(* IEC 61131-3 sources: daoli-st-library/DL_Process (part 61) *)

(* ---- FB_DL_BatchDosingControl.st ---- *)
(*==============================================================================
 * 组件名称 (Component)  : FB_DL_BatchDosingControl
 * 所属子库 (Sublibrary) : DL_Process
 * 当前版本 (Version)    : 1.0.1
 * 兼容性 (Platform)   : CODESYS 3.5 / TwinCAT 3 / 汇川 InoProShop / Machine Expert
 *                         仅依赖 Standard.library（TON / R_TRIG），零厂商方言
 * 分类     (Category)   : 工艺功能块（Function Block · 多原料单通道配料称重）
 * 功能简述 (Function)   : 多原料单通道自动配料称重控制器（单料批次相 Phase
 *                         语义）。三段给料顺控（快加→慢加→落定结算）+ 空中
 *                         落差自学习（误差/2 更新，防振荡）+ 超差 NG 判定 +
 *                         断流诊断。执行机构抽象为三离散输出（与给料机/闸门
 *                         类型解耦）；秤重量 LREAL→REAL 引脚注入（标定由称
 *                         重层完成）。Abort 优先级最高（CASE 首分支）。
 * 枚举归属 (Enum note)  : E_DL_DosingPhase 随本块同文件发布（公约 0.11 口径：
 *                         配套枚举与主块同文件，头注释注明归属）。
 * 公约遵循 (Convention) : 0.1/R23 显式批次启动沿驱动（无自动首扫初始化语义），
 *                         免首扫，无 bInit。
 *                         0.2/R21 bFault 显式排除信息级码；0.5/R7 全部实例主
 *                         体最前部无条件刷新；0.7/R15 断流/秤信号/参数故障锁
 *                         存仅复位路径清码；0.9 非有限值 fWeight 防御（自比
 *                         检测，故障级中止全断）；0.14 全部除法/浮点判等走
 *                         ABS 容差。
 *                         0.8 故障码段位 16#0005_xxxx（经 DL_Process
 *                         VERSION.md 码表核对，0005_0220~0223 / 0005_0114~0106
 *                         均未占用）：
 *                         【故障级】0005_0220 断流/堵料、0005_0221 秤信号无
 *                         效（非有限值）、0005_0223 配方参数非法、0005_0222
 *                         非法状态兜底；
 *                         【信息级】0005_0114 稳窗超时按当前值结算、0005_0115
 *                         补偿学习触限。
 * 红线自检 (Redline)    : R1 零全局变量表/外部变量引用 ✓｜R2 零物理 IO 地址 ✓
 *                         R3 纯 IEC 61131-3 ✓｜R4 非有限值中止全断/防振荡半
 *                         误差学习/限幅钳位 ✓
 *                         R5 全变量中英双语同行注释 ✓｜R6 ENUM+CASE+ELSE，Abort
 *                         首分支最高优先 ✓
 *                         R7 五实例（R_TRIG×3/TON×2）主体最前部无条件刷新 ✓
 *                         R8 全常量化 ✓
 * 设计要点 (Key notes)  : ① 截断点公式：慢加关断重量 = fSetpoint −
 *                           fInflightComp；fInflightComp 初值 0 → 首批必然过
 *                           冲 → 学习链收敛（首批预期在注释写明）；
 *                         ② 自学习更新：结算后 Error = fFinalWeight −
 *                           fSetpoint；bLearnEnable 时 fInflightComp +=
 *                           Error/2.0（半误差防振荡），钳位 ±fCompLimit，
 *                           触限置信息级 0005_0115；
 *                         ③ 稳窗判稳：tSettleWindow 内重量变化 <
 *                           fFlowDeadband 才结算；超窗未稳重试
 *                           DL_SETTLE_RETRY_MAX 次后按当前值结算 + 信息级；
 *                         ④ 断流诊断：给料相中 tFlowWatch 窗内重量变化 <
 *                           fFlowDeadband → 断流故障锁存（快加/慢加独立监
 *                           视计时重启）；
 *                         ⑤ 超差 NG 锁存 + 卸料输出禁止（NG 不得流入下工
 *                           序）；Abort 电平最高优先（CASE 首分支，立即关全
 *                           部输出）；
 *                         ⑥ 非有限值 fWeight → 批次中止故障级 0005_0221，
 *                           输出全断。
 * 偏离留档 (Deviation)  : 依 R11 头注释留档，共 1 条：
 *                         ① 新增故障码 0005_0223 配方参数非法：规格故障集未
 *                           覆盖 fSetpoint/fTolerance 非法值路径，编码时补
 *                           充登记（核对 DL_Process 码表未占用）。
 * 开源溯源 (Origin)     : 来源标签 lbp-batch-dosing / isa-88（RAW_NOTES_R7
 *                         S-10：ISA-88 批次相（Phase）语义与重力失重式/增
 *                         量式配料公开工程惯例——三段给料、空中落差补偿、
 *                         半误差学习（提取点②③⑤），公开技术资料，仅借鉴
 *                         语义域；状态机、学习与诊断实现、码位与引脚契约
 *                         100% 本库独立设计，clean-room 未复制源码）。
 * 验收向量 (Acceptance) :
 *   V1 三段给料逐拍：快加至 fSetpoint−fInflightComp 切慢加，同点关断进落定；
 *   V2 学习链 5 批收敛数值复算：首批过冲 Δ → 补偿 +Δ/2 → 逐批 Δ 减半；
 *   V3 补偿限幅：学习值触及 ±fCompLimit → 信息级 0005_0115；
 *   V4 断流：给料中 tFlowWatch 内重量变化 < fFlowDeadband → 0005_0220；
 *   V5 超差 NG + 卸料禁止：|误差| > fTolerance → eNg、bOutDischarge=FALSE；
 *   V6 中止优先级：任意相 bCmdAbort 电平 → 全输出断进 eAbort；
 *   V7 非有限值注入：fWeight=NaN → 0005_0221 输出全断。
 * 修订历史 (Revision)   :
 *   2026-11-15  v1.0.0  首版入库（Round 07 · DL_Process 配料称重件）
 *   2026-11-15  v1.0.1  终审修复 2 处：① _bSettleRestart/_bFlowRestart 单拍
 *                       重启标志永不自清 → 稳窗 TON 永久失效（eSettling 永
 *                       久挂起、判稳拍结算死锁）+ 断流诊断一次后失效（段 1
 *                       实例调用后自清，R24 同源范式）；② fTareOffset/
 *                       fInflightComp 缺 0.9 非数防御（NaN 扩散进净重/截
 *                       断点链路），新增 _fTareEff/_fCompEff 生效值
 *============================================================================*)

(*-----------------------------------------------------------------------------
 * 枚举: E_DL_DosingPhase（归属 FB_DL_BatchDosingControl，与其同文件）
 * 含义: 单料批次相离散状态。编号步长 10 留空位，eFault 取 99 保证排序末位
 *       （全库枚举编号惯例）。
 *----------------------------------------------------------------------------*)
TYPE E_DL_DosingPhase :
(
    eIdle     := 0,   // 空闲：等待批次启动 / Idle, awaiting batch start
    eCoarse   := 10,  // 快加：粗给料输出有效 / Coarse feed active
    eFine     := 20,  // 慢加：细给料输出有效 / Fine feed active
    eSettling := 30,  // 落定：稳窗判稳中 / Settling, stability window judging
    eDone     := 40,  // 完成：批次合格，卸料输出有效 / Done, batch OK, discharge active
    eNg       := 50,  // 超差：批次 NG 锁存，卸料禁止 / NG latched, discharge forbidden
    eAbort    := 60,  // 中止：Abort 电平保持中，全输出断 / Aborted, all outputs off
    eFault    := 99   // 故障锁存：断流/秤信号/参数非法/非法状态 / Latched fault
) UINT;
END_TYPE

FUNCTION_BLOCK FB_DL_BatchDosingControl
VAR_INPUT
    bCmdBatchStart : BOOL;              // 批次启动指令（Batch start），上升沿进入快加 / Batch start edge enters coarse feed
    bCmdAbort      : BOOL;              // 批次中止指令（Abort），电平生效，立即关全部输出 / Abort level, all outputs off immediately
    fWeight        : REAL;              // 秤实时重量（Live weight）[kg]，非有限值防御；标定由称重层完成 / Live weight [kg], non-finite defended, calibration upstream
    fTareOffset    : REAL := 0.0;       // 皮重偏移（Tare offset）[kg]，默认 0.0；净重 = fWeight − fTareOffset / Tare offset [kg], net = weight − tare
    fSetpoint      : REAL;              // 批次目标净重（Batch setpoint）[kg]，域 >0 / Batch setpoint [kg], > 0
    fSwitchCoarse  : REAL := 0.0;       // 快加切换点（Coarse-to-fine switch）[kg]，0=默认 85% 设定值（引脚覆盖语义见头注释）/ Coarse switch point, 0 = default 85% of setpoint
    fInflightComp  : REAL;              // 空中落差补偿（In-flight compensation）[kg]，学习值跨批次保持；上下限由 fCompLimit 钳位 / In-flight compensation [kg], learned value clamped by fCompLimit
    fCompLimit     : REAL := 0.0;       // 补偿学习限幅（Compensation limit）[kg]，0=默认 10% 设定值 / Compensation clamp, 0 = default 10% of setpoint
    bLearnEnable   : BOOL;              // 落差自学习使能（Learning enable），TRUE=每批结算后按误差/2 更新 / Learning enable, update by error/2 after each settle
    tSettleWindow  : TIME := T#1S;     // 落定稳窗（Settle window），默认 T#1S，域 500MS~5S 越界钳位 / Settle window, clamped 500MS..5S
    fTolerance     : REAL := 0.0;       // 批次公差（Batch tolerance）[kg]，0=默认 0.5% 设定值语义（引脚显式覆盖）/ Batch tolerance, 0 = default 0.5% of setpoint
    tFlowWatch     : TIME := T#10S;    // 断流监视窗（Flow watchdog），默认 T#10S；给料中重量变化率恒零超窗 → 断流 / Flow watchdog, constant-weight over window = no flow
    fFlowDeadband  : REAL := 0.05;     // 断流判据死区（Flow deadband）[kg]，默认 0.05；稳窗内重量变化 < 死区判断流 / Flow deadband [kg], change below deadband = no flow
    bReset         : BOOL;              // 上升沿复位故障（Reset edge）/ Rising edge resets fault
END_VAR
VAR_OUTPUT
    bOutCoarse    : BOOL;               // 快加输出（Coarse feed output），给料机/闸门快加速率 / Coarse feed output
    bOutFine      : BOOL;               // 慢加输出（Fine feed output）/ Fine feed output
    bOutDischarge : BOOL;               // 卸料输出（Discharge output），批次合格后放料 / Discharge output, opens after batch OK
    fNetWeight    : REAL;               // 当前净重（Net weight）[kg] / Current net weight [kg]
    fFinalWeight  : REAL;               // 上批次结算净重（Final weight）[kg]，落定后锁存 / Final settled weight [kg], latched after settle
    bBatchOk      : BOOL;               // 批次合格（Batch OK），|结算净重 − 设定值| ≤ 公差 / Batch OK verdict
    bFault        : BOOL;               // 故障标志（Fault flag），显式排除信息级 / Fault flag, info codes excluded
    uErrorId      : UDINT;              // 故障码（Error code），16#0005_xxxx 段，0=无故障 / Error code, family 16#0005_xxxx
END_VAR
VAR
    _ePhase        : E_DL_DosingPhase := E_DL_DosingPhase.eIdle; // 内部批次相（Internal dosing phase），属性只读 / Internal phase, read-only via property
    _bFaultLatch   : BOOL;              // 故障锁存标志（Fault latch flag），仅复位路径清除 / Fault latch, cleared only via reset path
    _uErrorIdInt   : UDINT;             // 内部故障级码寄存（Internal fault-level register）/ Internal fault-level register
    _uInfoCode     : UDINT;             // 本拍信息级码（Info code this cycle），瞬时型每拍重算 / Transient info code, recomputed each scan
    _bWeightValid  : BOOL;              // 秤信号有效（Weight signal valid，非有限值防御）/ Weight signal valid flag
    _fNetInt       : REAL;              // 内部净重（Internal net weight）[kg] / Internal net weight [kg]
    _fSetEff       : REAL;              // 防御后生效设定值（Sanitized setpoint）[kg] / Sanitized setpoint [kg]
    _fTolEff       : REAL;              // 防御后生效公差（Sanitized tolerance）[kg] / Sanitized tolerance [kg]
    _fSwitchEff    : REAL;              // 防御后生效快加切换点（Sanitized coarse switch）[kg] / Sanitized coarse switch [kg]
    _fCompLimEff   : REAL;              // 防御后生效补偿限幅（Sanitized compensation clamp）[kg] / Sanitized compensation clamp [kg]
    _fTareEff      : REAL;              // 防御后生效皮重偏移（Sanitized tare offset）[kg]，0.9 非数防御 / Sanitized tare offset [kg] (v1.0.1)
    _fCompEff      : REAL;              // 防御后生效落差补偿（Sanitized in-flight comp）[kg]，0.9 非数防御 / Sanitized in-flight comp [kg] (v1.0.1)
    _fCutCoarse    : REAL;              // 快加→慢加切换重量（Coarse-to-fine cut weight）[kg] / Coarse-to-fine cut weight [kg]
    _fCutFine      : REAL;              // 慢加关断重量（Fine cut weight）[kg]，= 设定值 − 落差补偿 / Fine cut weight [kg]
    _fSettleRef    : REAL;              // 稳窗基准重量（Settle reference weight）[kg] / Settle reference weight [kg]
    _nSettleRetry  : USINT;             // 稳窗重试计数（Settle retry counter）/ Settle retry counter
    _bSettleRestart: BOOL;              // 稳窗重启单拍（Settle restart one-shot）/ Settle restart one-shot
    _fFlowRef      : REAL;              // 断流监视基准重量（Flow-watch reference weight）[kg] / Flow-watch reference weight [kg]
    _bFlowRestart  : BOOL;              // 断流监视重启单拍（Flow-watch restart one-shot）/ Flow-watch restart one-shot
    _bBatchStartEdge : BOOL;            // 批次启动沿（Batch start edge this scan）/ Batch start edge this scan
    _fbTrigStart   : R_TRIG;            // 批次启动沿检测（Batch start edge detector）/ Batch start edge detector
    _fbTrigReset   : R_TRIG;            // 复位沿检测（Reset edge detector）/ Reset edge detector
    _fbTrigAbort   : R_TRIG;            // 中止沿检测（Abort edge detector），沿置中止态（电平保持由段内判定）/ Abort edge detector
    _fbTonSettle   : TON;               // 落定稳窗定时器（Settle window timer）/ Settle window timer
    _fbTonFlow     : TON;               // 断流监视窗定时器（Flow watchdog timer）/ Flow watchdog timer
END_VAR
VAR CONSTANT
    DL_COARSE_FRAC    : REAL := 0.85;   // 快加切换默认比例（Coarse switch default fraction of setpoint）/ Coarse switch default fraction
    DL_COMP_FRAC      : REAL := 0.10;   // 补偿限幅默认比例（Compensation clamp default fraction）/ Compensation clamp default fraction
    DL_TOL_FRAC       : REAL := 0.005;  // 公差默认比例（Tolerance default fraction of setpoint）/ Tolerance default fraction
    DL_LEARN_DIV      : REAL := 2.0;    // 学习半误差除数（Learning half-error divisor），防振荡 / Learning half-error divisor, anti-oscillation
    DL_SETTLE_WIN_MIN : TIME := T#500MS; // 稳窗下限（Settle window lower clamp）/ Settle window lower clamp
    DL_SETTLE_WIN_MAX : TIME := T#5S;   // 稳窗上限（Settle window upper clamp）/ Settle window upper clamp
    DL_SETTLE_RETRY_MAX : USINT := 3;   // 稳窗重试上限（Settle retry max），超限按当前值结算 / Settle retry max, settle as-is beyond
    DL_REAL_EPS       : REAL := 1.0E-6; // 浮点防零容差（Float divide-guard epsilon）/ Float divide-guard epsilon
END_VAR

// ============================================================================
// 段 1｜实例无条件周期刷新（R7/0.5：严禁置于 IF/CASE 分支内）
//      Unconditional per-cycle refresh of all instances (R7/0.5)
// ============================================================================
_fbTrigStart(CLK := bCmdBatchStart);
_fbTrigReset(CLK := bReset);
_fbTrigAbort(CLK := bCmdAbort);
_bBatchStartEdge := _fbTrigStart.Q;   // 本拍启动沿（Start edge this scan）
_fbTonSettle(IN := (_ePhase = E_DL_DosingPhase.eSettling) AND (NOT _bSettleRestart) AND (NOT _bFaultLatch), PT := tSettleWindow); // 稳窗（Settle window）
_fbTonFlow(IN := ((_ePhase = E_DL_DosingPhase.eCoarse) OR (_ePhase = E_DL_DosingPhase.eFine))
           AND (NOT _bFlowRestart) AND (NOT _bFaultLatch), PT := tFlowWatch); // 断流监视窗（Flow watchdog）
// R24 同源范式：单拍重启标志在实例调用之后自清（v1.0.1 修复：原永不自清 →
// 稳窗 TON 永久失效（eSettling 永久挂起、判稳拍结算死锁）+ 断流诊断一次后
// 永久失效）/ One-shot restart flags self-cleared AFTER the instance calls
// (v1.0.1 fix: flags were never cleared, permanently disabling both timers)
_bSettleRestart := FALSE;         // 稳窗重启单拍自清（Settle restart flag self-cleared）
_bFlowRestart := FALSE;           // 断流监视重启单拍自清（Flow restart flag self-cleared）

// ============================================================================
// 段 2｜秤信号防御（0.9）+ 信息级预清零 + 复位路径（R15）
//      Weight sanitation (0.9) + info preset + reset path (R15)
// ============================================================================
_uInfoCode := 0;                  // 信息级瞬时型每拍重算（Transient info recomputed each scan）

IF fWeight <> fWeight THEN        // 非数自比检测（NaN self-compare）
    _bWeightValid := FALSE;       // 秤信号无效（Weight invalid）
    IF _bFaultLatch = FALSE THEN
        _bFaultLatch := TRUE;     // 秤信号无效故障锁存（Invalid weight latch）
        _uErrorIdInt := 16#0005_0221; // 0005_0221 秤信号无效【故障级】/ Invalid weight signal, fault level
        _ePhase := E_DL_DosingPhase.eFault; // 批次中止进故障态（Batch aborted to fault）
    END_IF
ELSE
    _bWeightValid := TRUE;        // 秤信号有效（Weight valid）
    _fNetInt := fWeight - _fTareEff; // 净重计算（皮重经 0.9 非数防御生效值，v1.0.1）/ Net weight with sanitized tare (v1.0.1)
END_IF
fNetWeight := _fNetInt;           // 净重出口（Net weight outlet）

IF _fbTrigReset.Q THEN
    _bFaultLatch := FALSE;        // 故障锁存解除（Fault latch released）
    _uErrorIdInt := 16#0000_0000; // 故障码清零（Fault code cleared）
    IF _ePhase = E_DL_DosingPhase.eFault THEN
        _ePhase := E_DL_DosingPhase.eIdle; // 故障复位回空闲（Fault reset to idle）
    END_IF
END_IF

// ============================================================================
// 段 3｜参数防御（启动时校验配方，0.9 + 域防御）
//      Recipe parameter sanitation at batch start (0.9 + domain guards)
// ============================================================================
IF fSetpoint <> fSetpoint THEN    // 设定值非数（Setpoint NaN）
    _fSetEff := 0.0;              // 非法设定占位（Invalid placeholder）
ELSIF fSetpoint <= DL_REAL_EPS THEN
    _fSetEff := 0.0;              // 非正设定占位（Non-positive placeholder）
ELSE
    _fSetEff := fSetpoint;        // 生效设定（Effective setpoint）
END_IF

IF fTolerance <> fTolerance THEN  // 公差非数（Tolerance NaN）
    _fTolEff := _fSetEff * DL_TOL_FRAC; // 回落默认比例（Default fraction fallback）
ELSIF fTolerance <= 0.0 THEN
    _fTolEff := _fSetEff * DL_TOL_FRAC; // 非正回落默认（Non-positive falls back）
ELSE
    _fTolEff := fTolerance;       // 生效公差（Effective tolerance）
END_IF

IF fSwitchCoarse <> fSwitchCoarse THEN // 切换点非数（Switch NaN）
    _fSwitchEff := _fSetEff * DL_COARSE_FRAC; // 回落默认比例（Default fraction fallback）
ELSIF fSwitchCoarse <= 0.0 THEN
    _fSwitchEff := _fSetEff * DL_COARSE_FRAC; // 零值=默认 85% 设定值（Zero = default 85%）
ELSE
    _fSwitchEff := fSwitchCoarse; // 引脚覆盖生效（Pin override effective）
END_IF

IF fCompLimit <> fCompLimit THEN  // 限幅非数（Clamp NaN）
    _fCompLimEff := _fSetEff * DL_COMP_FRAC; // 回落默认比例（Default fraction fallback）
ELSIF fCompLimit <= 0.0 THEN
    _fCompLimEff := _fSetEff * DL_COMP_FRAC; // 零值=默认 10% 设定值（Zero = default 10%）
ELSE
    _fCompLimEff := fCompLimit;   // 生效限幅（Effective clamp）
END_IF

// 0.9 非数防御补齐（v1.0.1）：皮重偏移与落差补偿为 REAL 输入，非数自比后
// 取生效值，杜绝 NaN 扩散进净重/截断点链路
// 0.9 NaN defense completed (v1.0.1) for tare offset and in-flight compensation
IF fTareOffset <> fTareOffset THEN // 皮重非数（Tare NaN）
    _fTareEff := 0.0;             // 回落零皮重（Fallback zero tare）
ELSE
    _fTareEff := fTareOffset;     // 生效皮重（Effective tare）
END_IF
IF fInflightComp <> fInflightComp THEN // 落差补偿非数（In-flight comp NaN）
    _fCompEff := 0.0;             // 回落零补偿（首批过冲语义，学习链重建）/ Fallback zero comp
ELSE
    _fCompEff := fInflightComp;   // 生效补偿（Effective compensation）
END_IF

// ============================================================================
// 段 4｜主批次相状态机（ENUM + CASE + ELSE 兜底；Abort 首分支最高优先）
//      Main dosing phase machine (Abort first-branch top priority, ELSE fallback)
// ============================================================================
IF bCmdAbort THEN
    // Abort 电平最高优先：立即关全部输出进中止态（Abort level top priority）
    _ePhase := E_DL_DosingPhase.eAbort; // 进中止态（To aborted state）
ELSE
    CASE _ePhase OF

        E_DL_DosingPhase.eIdle: // 空闲态：等待启动沿
            IF _bBatchStartEdge AND (NOT _bFaultLatch) THEN
                IF _fSetEff <= DL_REAL_EPS THEN
                    _bFaultLatch := TRUE;           // 配方参数非法锁存（Invalid recipe latch）
                    _uErrorIdInt := 16#0005_0223;   // 0005_0223 配方参数非法【故障级】/ Invalid recipe parameters, fault level
                    _ePhase := E_DL_DosingPhase.eFault;
                ELSE
                    _fCutCoarse := _fSwitchEff;                     // 快加切换点（Coarse cut point）
                    _fCutFine := _fSetEff - _fCompEff;              // 慢加关断重量 = 设定值 − 落差补偿（截断点公式，生效值）/ Fine cut = setpoint − sanitized comp
                    fFinalWeight := 0.0;                            // 上批结果清位（Final weight cleared）
                    bBatchOk := FALSE;                              // 合格判定清位（OK verdict cleared）
                    _nSettleRetry := 0;                             // 稳窗重试清零（Retry cleared）
                    _fSettleRef := _fNetInt;                        // 稳窗基准初始化（Settle reference init）
                    _fFlowRef := _fNetInt;                          // 断流基准初始化（Flow reference init）
                    _ePhase := E_DL_DosingPhase.eCoarse;            // 进入快加（To coarse feed）
                END_IF
            END_IF

        E_DL_DosingPhase.eCoarse: // 快加态：粗给料至切换点
            IF _fNetInt >= _fCutCoarse THEN
                _ePhase := E_DL_DosingPhase.eFine; // 切慢加（To fine feed）
                _fFlowRef := _fNetInt;             // 断流基准重置（Flow reference reset）
            END_IF

        E_DL_DosingPhase.eFine: // 慢加态：细给料至截断点
            IF _fNetInt >= _fCutFine THEN
                _ePhase := E_DL_DosingPhase.eSettling; // 关断进落定（Cut to settling）
                _fSettleRef := _fNetInt;               // 稳窗基准重置（Settle reference reset）
            END_IF

        E_DL_DosingPhase.eSettling: // 落定态：稳窗判稳，判稳即一次性结算+学习
            IF _fbTonSettle.Q THEN
                IF ABS(_fNetInt - _fSettleRef) < fFlowDeadband THEN
                    // —— 一次性结算（仅判稳拍执行）：锁存结果 + NG 判定 + 学习 ——
                    //     One-shot settlement on the settled scan: result latch, NG verdict, learning
                    fFinalWeight := _fNetInt;   // 结算净重锁存（Final weight latched）
                    bBatchOk := ABS(fFinalWeight - _fSetEff) <= _fTolEff; // 公差判定（Tolerance verdict）
                    IF bLearnEnable THEN
                        fInflightComp := fInflightComp + (fFinalWeight - _fSetEff) / DL_LEARN_DIV; // 误差/2 学习（半误差防振荡）/ Half-error learning, anti-oscillation
                        IF fInflightComp > _fCompLimEff THEN
                            fInflightComp := _fCompLimEff;  // 正向限幅（Positive clamp）
                            _uInfoCode := 16#0005_0115;     // 0005_0115 补偿学习触限【信息级】/ Learning clamp hit, info level
                        ELSIF fInflightComp < (-_fCompLimEff) THEN
                            fInflightComp := -_fCompLimEff; // 负向限幅（Negative clamp）
                            _uInfoCode := 16#0005_0115;     // 0005_0115 补偿学习触限【信息级】/ Learning clamp hit, info level
                        END_IF
                    END_IF
                    IF bBatchOk THEN
                        _ePhase := E_DL_DosingPhase.eDone;  // 合格进完成态（OK to done）
                    ELSE
                        _ePhase := E_DL_DosingPhase.eNg;    // 超差进 NG 锁存态（Out of tolerance to NG）
                    END_IF
                ELSE
                    _nSettleRetry := _nSettleRetry + 1; // 未稳重试（Retry when unstable）
                    IF _nSettleRetry >= DL_SETTLE_RETRY_MAX THEN
                        _uInfoCode := 16#0005_0114;     // 0005_0114 稳窗超时按当前值结算【信息级】/ Settle timeout, settle as-is, info level
                        fFinalWeight := _fNetInt;       // 按当前值结算锁存（Settle as-is latch）
                        bBatchOk := ABS(fFinalWeight - _fSetEff) <= _fTolEff; // 公差判定（Tolerance verdict）
                        IF bBatchOk THEN
                            _ePhase := E_DL_DosingPhase.eDone;
                        ELSE
                            _ePhase := E_DL_DosingPhase.eNg;
                        END_IF
                    ELSE
                        _fSettleRef := _fNetInt;        // 重置稳窗基准（Reset settle reference）
                        _bSettleRestart := TRUE;        // 稳窗重启单拍（Restart window one-shot）
                    END_IF
                END_IF
            END_IF

        E_DL_DosingPhase.eDone: // 完成态：卸料保持，等待新批次启动
            IF _bBatchStartEdge AND (NOT _bFaultLatch) THEN
                IF _fSetEff <= DL_REAL_EPS THEN
                    _bFaultLatch := TRUE;               // 配方参数非法锁存（Invalid recipe latch）
                    _uErrorIdInt := 16#0005_0223;       // 0005_0223 配方参数非法【故障级】/ Invalid recipe, fault level
                    _ePhase := E_DL_DosingPhase.eFault;
                ELSE
                    _fCutCoarse := _fSwitchEff;         // 快加切换点（Coarse cut point）
                    _fCutFine := _fSetEff - _fCompEff;  // 截断点更新（Fine cut update, sanitized comp）
                    fFinalWeight := 0.0;                // 上批结果清位（Final weight cleared）
                    bBatchOk := FALSE;                  // 合格判定清位（OK verdict cleared）
                    _nSettleRetry := 0;                 // 稳窗重试清零（Retry cleared）
                    _fSettleRef := _fNetInt;            // 稳窗基准初始化（Settle reference init）
                    _fFlowRef := _fNetInt;              // 断流基准初始化（Flow reference init）
                    _ePhase := E_DL_DosingPhase.eCoarse; // 进入快加（To coarse feed）
                END_IF
            END_IF

        E_DL_DosingPhase.eNg: // 超差态：卸料禁止，等待新批次启动或 Abort
            IF _bBatchStartEdge AND (NOT _bFaultLatch) THEN
                IF _fSetEff <= DL_REAL_EPS THEN
                    _bFaultLatch := TRUE;               // 配方参数非法锁存（Invalid recipe latch）
                    _uErrorIdInt := 16#0005_0223;       // 0005_0223 配方参数非法【故障级】/ Invalid recipe, fault level
                    _ePhase := E_DL_DosingPhase.eFault;
                ELSE
                    _fCutCoarse := _fSwitchEff;         // 快加切换点（Coarse cut point）
                    _fCutFine := _fSetEff - _fCompEff;  // 截断点更新（Fine cut update, sanitized comp）
                    fFinalWeight := 0.0;                // 上批结果清位（Final weight cleared）
                    bBatchOk := FALSE;                  // 合格判定清位（OK verdict cleared）
                    _nSettleRetry := 0;                 // 稳窗重试清零（Retry cleared）
                    _fSettleRef := _fNetInt;            // 稳窗基准初始化（Settle reference init）
                    _fFlowRef := _fNetInt;              // 断流基准初始化（Flow reference init）
                    _ePhase := E_DL_DosingPhase.eCoarse; // 重开新批（New batch from coarse）
                END_IF
            END_IF

        E_DL_DosingPhase.eAbort: // 中止态：Abort 电平撤销后回空闲
            IF NOT bCmdAbort THEN
                _ePhase := E_DL_DosingPhase.eIdle; // 电平撤销回空闲（Level dropped, back to idle）
            END_IF

        E_DL_DosingPhase.eFault: // 故障锁存态：复位路径见段 2
            // 等待复位（Await reset）

        ELSE
            // 非法状态兜底：任何越界枚举值强制锁存故障（Illegal state fallback）
            _bFaultLatch := TRUE;           // 故障锁存（Fault latch）
            _uErrorIdInt := 16#0005_0222;   // 0005_0222 非法状态兜底【故障级】/ Illegal state, fault level
            _ePhase := E_DL_DosingPhase.eFault;
    END_CASE
END_IF

// ============================================================================
// 段 5｜输出推导 + 断流诊断 + 输出全断出口断言
//      Output derivation + no-flow diagnosis + all-off exit assertion
// ============================================================================
bOutCoarse := (_ePhase = E_DL_DosingPhase.eCoarse) AND _bWeightValid AND (NOT _bFaultLatch); // 快加输出派生（Coarse derived form）
bOutFine := (_ePhase = E_DL_DosingPhase.eFine) AND _bWeightValid AND (NOT _bFaultLatch);     // 慢加输出派生（Fine derived form）
bOutDischarge := (_ePhase = E_DL_DosingPhase.eDone) AND bBatchOk AND (NOT _bFaultLatch);     // 卸料输出派生（NG/Abort/故障恒断，出口断言）/ Discharge derived, off on NG/abort/fault

// 断流诊断：监视窗到且给料相中重量未前进死区 → 断流锁存（快加/慢加独立重置基准）
// No-flow diagnosis: watchdog expired in feed phases without weight advance
IF _fbTonFlow.Q THEN
    IF ABS(_fNetInt - _fFlowRef) < fFlowDeadband THEN
        _bFaultLatch := TRUE;         // 断流故障锁存（No-flow latch）
        _uErrorIdInt := 16#0005_0220; // 0005_0220 断流/堵料【故障级】/ No flow or bridging, fault level
        _ePhase := E_DL_DosingPhase.eFault;
    ELSE
        _fFlowRef := _fNetInt;        // 基准前移（Reference advanced）
        _bFlowRestart := TRUE;        // 监视窗重启单拍（Watchdog restart one-shot）
    END_IF
END_IF

(*------------------------------------------------------------------------------
 * 属性: ePhase（GET）—— 当前批次相只读视图（Phase 语义对外镜像）。
 *      Property ePhase (GET) - read-only dosing phase view.
 *------------------------------------------------------------------------------*)
PROPERTY ePhase : E_DL_DosingPhase
ePhase := _ePhase;                // 返回内部批次相（Return internal phase）
END_PROPERTY

(*------------------------------------------------------------------------------
 * 属性: bFault（GET）—— 故障锁存指示（信息级码不置本位，0.2 公约）。
 *      Property bFault (GET) - fault latch indicator, info codes excluded.
 *------------------------------------------------------------------------------*)
PROPERTY bFault : BOOL
bFault := _bFaultLatch OR (_ePhase = E_DL_DosingPhase.eFault); // 显式排除信息级派生式（Derived form excluding info codes）
END_PROPERTY

(*------------------------------------------------------------------------------
 * 属性: uErrorId（GET）—— 末次故障码（故障级优先，无故障时透出本拍信息级
 *         码，0.2/0.15 公约）。
 *      Property uErrorId (GET) - last error code (fault priority, info shown otherwise).
 *------------------------------------------------------------------------------*)
PROPERTY uErrorId : UDINT
IF (_uErrorIdInt <> 0) OR (_ePhase = E_DL_DosingPhase.eFault) THEN
    uErrorId := _uErrorIdInt;     // 故障级码优先透出（Fault-level priority）
ELSE
    uErrorId := _uInfoCode;       // 无故障时透出本拍信息级码（Transient info code）
END_IF
END_PROPERTY
END_FUNCTION_BLOCK

(* ---- FB_DL_BatchPhaseBase.st ---- *)
(*==============================================================================
 * 组件名称 (Component)  : FB_DL_BatchPhaseBase
 * 所属子库 (Sublibrary) : DL_Process
 * 当前版本 (Version)    : 1.0.1
 * 组件分类 (Category)   : 功能块（FUNCTION_BLOCK）· 批次工艺 · 相状态机底座
 * 兼容性   (Platform)   : CODESYS 3.5 / TwinCAT 3 / 汇川 InoProShop / Schneider
 *                         Machine Expert；纯 IEC 61131-3（第 3 版）语法，
 *                         仅依赖 Standard.library（R_TRIG / TON）
 * 功能描述 (Function)   : ISA-88 批次相（Phase）的标准状态机底座：提供相状态迁移、
 *                         相内步骤推进、暂停与恢复、停止与中止四类命令的语义裁决，
 *                         以及相净运行时间累计。具体工艺动作不在本件内实现，由调用方
 *                         按「步骤执行请求」外置实现，完成或失败再回送反馈。
 * 分层声明 (Layering)   : ① 本件不实现任何工艺动作（投料、升温、搅拌、清洗的开阀与
 *                         设定值下发都在调用方），也不定义配方与流程结构（配方、程序、
 *                         单元编排属上层，另立件）；
 *                         ② 本件不驱动任何设备，不读写工艺参数，只裁决状态与命令；
 *                         ③ 步骤动作外置带来一个必须遵守的约定：收到步骤执行请求后，
 *                         调用方要自行记住「当前步已启动」，再用完成或失败反馈应答。
 * 语义要点 (Semantics)  :
 *   ① 命令优先级严格为 中止 高于 停止 高于 暂停 高于 恢复 高于 启动；同拍多命令时高
 *      优先者胜，低优先者直接丢弃且**不排队**——排队会让操作员的「停止」在几拍之后
 *      突然生效，属高危行为。
 *   ② 暂停只在步骤边界生效：暂停请求先登记，等当前步骤的完成反馈被消费、或步骤请求
 *      尚未发出时才真正进入暂停。**绝不在动作执行中途切断**，这是相语义的核心，也是
 *      现场「暂停后物料半投」事故的根因。
 *   ③ 恢复不重头：恢复时步骤号保持不变，重新发当前步骤的执行请求，从该步继续。
 *   ④ 已终止态（完成、已停、已中止）不接受启动与中止命令，只接受复位。
 *   ⑤ 掉使能时冻结状态与全部输出、不清零——批次报表需要看到最后相状态。
 * 计时口径 (Elapsed)    : 相运行累计时间只在执行相累加，暂停相与其余相不计入，故该值
 *                         即「相净运行时间」，MES 用它算相耗时与产能。
 * 开源溯源 (Origin)     : 来源标签 isa88-batch。原创实现（参考 ISA-88 与 IEC 61512 公开的
 *                         相状态模型：空闲、执行、收尾、完成、暂停请求、已暂停、恢复中、
 *                         停止中、已停、中止中、已中止的状态集合，以及「暂停在步骤边界
 *                         生效」「恢复不重头」两条语义）。ISA-88 为公开规范而非代码，
 *                         无代码复制问题；成员编号、状态机实现、超时策略、单拍请求语义、
 *                         计时口径与全部码位 100% 本库独立设计，clean-room 实现。
 * 依赖     (Depends)    : 无 DL_ 内部依赖；Standard.library: R_TRIG / TON
 * 故障码表 (Error codes):
 *   16#0005_0104【信息级】相内步骤数越界已钳到 1 至 32
 *   16#0005_0105【信息级】同拍多命令，低优先命令已丢弃（不排队）
 *   16#0005_0106【信息级】从暂停恢复，步骤号不重置
 *   16#0005_0107【信息级】单步或暂停超时监控被关闭（参数为 0）
 *   16#0005_0203【故障级】单步超时，相中止（锁存）
 *   16#0005_0204【故障级】步骤失败反馈，相中止（锁存，与完成反馈同拍时失败优先）
 *   16#0005_0205【故障级】暂停超时，相中止（锁存）
 *   16#0005_0206【故障级】非法状态兜底（锁存，直接进已中止，不回空闲）
 * 码位占用 (Slot)       : 信息级 0104 / 0105 / 0106 / 0107；故障级 0203 / 0204 / 0205 / 0206。
 *                         全部落在 R12 本件分配块内，无跨块借用、无段外哨兵值。
 * 拍序纪律 (Cycle order) :
 *   ① eState     ：段 7 状态机（唯一位移点），段 8 复位分支是唯一回空闲点
 *   ② nStep      ：进入执行相置 1、步骤推进加 1、复位清零，三处互斥
 *   ③ bStepAcked ：消费一次完成反馈即置位，反馈电平落下即清零（R34 状态量生命周期）
 *   ④ uErrorId   ：段 9 单一优先级链，全拍只写一次
 * 验收向量 (Acceptance) :
 *   V1 三步走完：步骤数 3，启动后每拍给一次完成反馈 → 依次执行 1、2、3 步，
 *      第三步完成进收尾，收尾完成进完成相，完成标志为真
 *   V2 步骤边界暂停：第 2 步执行中给暂停 → 先进暂停请求相，该步完成反馈到达后才进
 *      已暂停，此时不再发步骤请求；恢复后回执行相且步骤号仍为 2
 *   V3 中止与复位：已暂停时给中止 → 中止相发出中止动作单拍 → 已中止；复位回空闲、
 *      步骤号归零、完成标志清零
 *   V4 单步超时：单步超时 2 秒、步骤数 1、启动后不给完成反馈 → 2 秒后进中止、
 *      故障位置位、码 0203
 *   V5 失败优先：完成反馈与失败反馈同拍 → 进中止、码 0204
 * 偏离留档 (Deviation)  :
 *   ① 规格内部变量清单列有循环守卫量，本件无循环（步骤数固定上限、无数组遍历），
 *      故不声明，避免声明不用的死变量。
 *   ② 新增「步骤完成反馈」的上升沿实例（规格清单未列）。理由：若只靠电平消费，完成
 *      反馈常高时新步骤的完成永远等不到下降沿，会把相卡死在执行相（R34 只置不销）。
 *      上升沿实例与电平标志双保险，仍保留步骤已消费标志。
 *   ③ 规格写「恢复时把步骤已消费标志置真」，照写会把恢复后本步的完成反馈永久屏蔽，
 *      故按语义改为置假（恢复后重新等待本步的完成反馈），并写进头注释。
 *   ④ 停止请求在步骤边界生效后，收尾完成由调用方再给一次完成反馈；若收尾无反馈，
 *      单步超时会把相带进中止（宁停不悬）。
 * 修订历史 (Revision)   :
 *   2026-11-15  v1.0.0  首版落盘（R12 · 泳道 C · 批次相状态底座）
 *   2026-11-15  v1.0.1  终审修复两处：
 *                       ① 单步超时被实现成「相内累计超时」——监控定时器的输入在执行、收尾、
 *                       停止三相间持续为真，步骤推进时从不断输入，ET 跨步累加；3 步各 30 s、
 *                       超时 60 s 的合规批次会在第 3 步被误判 0203 中止。改为步骤边界断输入
 *                       一拍（bStepWatchBreak），超时按步重计时。
 *                       ② bStart 引脚注释原写「空闲与已终止态受理」，与实现（仅空闲受理、
 *                       终止态须先复位）不符，按实现更正注释
 *============================================================================*)

(*------------------------------------------------------------------------------
 * 枚举: E_DL_BatchPhaseState（相状态，归属本功能块并同文件发布）
 *       Phase state enumeration following the published ISA-88 phase model
 *       编号约定：0 起跳、步长 10，已中止取 99 保证排序末位
 *-----------------------------------------------------------------------------*)
TYPE E_DL_BatchPhaseState :
(
    eIdle       := 0,   // 空闲：等待启动，输出全复位 / Idle, waiting for the start command
    eRunning    := 10,  // 执行：按步骤号推进相内步骤 / Running, stepping through the phase
    eCompleting := 20,  // 收尾：最后一步已完成，等待收尾动作反馈 / Completing, waiting for the clean-up feedback
    eComplete   := 30,  // 完成：正常完成，保持到复位 / Complete, held until reset
    eHolding    := 40,  // 暂停请求：已受理，等步骤边界 / Holding, the hold request is accepted and pending a boundary
    eHeld       := 50,  // 已暂停：不再推进、不发步骤请求 / Held, no step request is issued
    eRestarting := 60,  // 恢复中：重发当前步骤请求，不重头 / Restarting, the current step is re-requested
    eStopping   := 70,  // 停止中：当前步骤收尾 / Stopping, the current step is being wrapped up
    eStopped    := 80,  // 已停：保持到复位 / Stopped, held until reset
    eAborting   := 90,  // 中止中：发出中止动作单拍 / Aborting, a one-scan abort request is issued
    eAborted    := 99   // 已中止：保持到复位 / Aborted, held until reset
);
END_TYPE

FUNCTION_BLOCK FB_DL_BatchPhaseBase
VAR_INPUT
    bEnable      : BOOL;                           // 使能，FALSE 时冻结状态与输出且不清零 [-] / Enable, freezes the phase without clearing it
    bStart       : BOOL;                           // 启动相，上升沿有效，仅空闲态受理（已终止态须先复位）[-] / Rising edge starts the phase in idle only, terminal states need a reset first
    bHold        : BOOL;                           // 请求暂停，上升沿有效，在步骤边界生效 [-] / Rising edge requests a hold at a step boundary
    bRestart     : BOOL;                           // 从已暂停恢复，上升沿有效，继续当前步骤 [-] / Rising edge resumes the current step
    bStop        : BOOL;                           // 请求停止，上升沿有效，在当前步骤完成后停 [-] / Rising edge requests a controlled stop
    bAbort       : BOOL;                           // 请求中止，上升沿有效，立即跳出步骤 [-] / Rising edge aborts immediately
    bReset       : BOOL;                           // 复位，上升沿有效，从已终止态回空闲 [-] / Rising edge returns the phase to idle
    bStepDone    : BOOL;                           // 步骤完成反馈（相内动作成功）[-] / Step completion feedback
    bStepFail    : BOOL;                           // 步骤失败反馈（相内动作失败）[-] / Step failure feedback
    nStepCount   : INT := 1;                       // 相内步骤数 [步]，有效域 1 到 32 / Steps in the phase, one to thirty-two
    tStepTimeout : TIME := T#60S;                  // 单步超时 [毫秒]，0 表示不监控 / Per-step timeout, zero disables the watchdog
    tHoldTimeout : TIME := T#600S;                 // 暂停超时 [毫秒]，0 表示不监控 / Hold timeout, zero disables the watchdog
END_VAR
VAR_OUTPUT
    ePhase       : E_DL_BatchPhaseState;           // 相状态，对外唯一状态出口 [-] / Phase state, the single state outlet
    nStepNo      : INT;                            // 当前步骤号，1 起，0 表示未进入 [步] / Current step number, zero before the first step
    bPhaseActive : BOOL;                           // 相处于活动族（执行、暂停族、收尾、停止、中止中）[-] / Phase is active
    bPhaseComplete : BOOL;                         // 相正常完成（完成相保持）[-] / Phase completed normally
    bRequestStep : BOOL;                           // 单拍：请执行当前步的动作 [-] / One-scan request to execute the current step
    bRequestAbort: BOOL;                           // 单拍：请执行中止动作 [-] / One-scan request to run the abort action
    uPhaseElapsed: UDINT;                          // 相净运行累计时间（不含暂停）[秒] / Accumulated running seconds excluding held time
    bError       : BOOL;                           // 故障级锁存，仅 0203 至 0206 置位 [-] / Latched fault, only fault level codes set it
    uErrorId     : UDINT;                          // 事件码，0 表示无事件 [代码] / Event code, zero means none
END_VAR
VAR
    fbTrigStart  : R_TRIG;                         // 启动沿检测，主周期无条件刷新 [-] / Start edge detector, refreshed unconditionally
    fbTrigHold   : R_TRIG;                         // 暂停沿检测，主周期无条件刷新 [-] / Hold edge detector, refreshed unconditionally
    fbTrigRestart: R_TRIG;                         // 恢复沿检测，主周期无条件刷新 [-] / Restart edge detector, refreshed unconditionally
    fbTrigStop   : R_TRIG;                         // 停止沿检测，主周期无条件刷新 [-] / Stop edge detector, refreshed unconditionally
    fbTrigAbort  : R_TRIG;                         // 中止沿检测，主周期无条件刷新 [-] / Abort edge detector, refreshed unconditionally
    fbTrigReset  : R_TRIG;                         // 复位沿检测，主周期无条件刷新 [-] / Reset edge detector, refreshed unconditionally
    fbTrigStepDone : R_TRIG;                       // 步骤完成上升沿，防电平常高时漏推进 [-] / Step completion rising edge
    fbStepWatch  : TON;                            // 单步超时监控，主周期无条件刷新 / Per-step watchdog, refreshed unconditionally
    fbHoldWatch  : TON;                            // 暂停超时监控，主周期无条件刷新 / Hold watchdog, refreshed unconditionally
    fbSecBase    : TON;                            // 一秒基准定时器，到点自复位 / One second base timer, self restarting
    bStepWatchBreak : BOOL;                        // 单步超时断输入一拍（步骤边界重计时）[-] / One-scan break of the step watchdog at a step boundary
    eState       : E_DL_BatchPhaseState := E_DL_BatchPhaseState.eIdle; // 内部相状态，对外经 ePhase 输出 [-] / Internal state exported as ePhase
    bInit        : BOOL := FALSE;                  // 首扫标志，初值 FALSE，判据取非 [-] / First-scan flag initialised FALSE
    bFaultLatch  : BOOL;                           // 故障锁存，仅复位分支清除 [-] / Fault latch, cleared by the reset path only
    uErrInt      : UDINT;                          // 故障级码寄存，锁存型 [代码] / Latched fault level code register
    uInfoCode    : UDINT;                          // 本拍信息级码，每拍重算 [代码] / Info level code recomputed every scan
    nStep        : INT;                            // 当前步骤号 [步]，0 表示未进入 / Current step number, zero before the first step
    nStepUse     : INT := 1;                       // 生效步骤数 [步]，钳位后 / Effective step count after clamping
    bStepIssued  : BOOL;                           // 本步执行请求已发出 [-] / Step request issued flag
    bStepAcked   : BOOL;                           // 本步完成反馈已被消费（防一步多次完成）[-] / Step completion consumed flag
    bHoldArmed   : BOOL;                           // 暂停请求已登记、待步骤边界生效 [-] / Hold armed, pending a step boundary
    bStopArmed   : BOOL;                           // 停止请求已登记 [-] / Stop armed
    bCmdStart    : BOOL;                           // 本拍生效的启动命令 [-] / Effective start command of this scan
    bCmdHold     : BOOL;                           // 本拍生效的暂停命令 [-] / Effective hold command of this scan
    bCmdRestart  : BOOL;                           // 本拍生效的恢复命令 [-] / Effective restart command of this scan
    bCmdStop     : BOOL;                           // 本拍生效的停止命令 [-] / Effective stop command of this scan
    bCmdAbort    : BOOL;                           // 本拍生效的中止命令 [-] / Effective abort command of this scan
    bCmdReset    : BOOL;                           // 本拍生效的复位命令 [-] / Effective reset command of this scan
    bCmdDropped  : BOOL;                           // 本拍存在被丢弃的低优先命令 [-] / A low priority command was dropped this scan
    bStepMon     : BOOL;                           // 单步超时监控启用 [-] / Step watchdog enabled
    bHoldMon     : BOOL;                           // 暂停超时监控启用 [-] / Hold watchdog enabled
    tStepUse     : TIME := T#60S;                  // 生效单步超时 [毫秒] / Effective step timeout
    tHoldUse     : TIME := T#600S;                 // 生效暂停超时 [毫秒] / Effective hold timeout
    bStepTo      : BOOL;                           // 单步超时到点 [-] / Step timeout reached
    bHoldTo      : BOOL;                           // 暂停超时到点 [-] / Hold timeout reached
    bSecTick     : BOOL;                           // 一秒脉冲 [-] / One second tick
    bSecDone     : BOOL;                           // 秒基准定时器到点电平，用于自复位 [-] / Second base elapsed level used for the self restart
    uElapsed     : UDINT;                          // 相净运行秒累计 [秒] / Accumulated running seconds
END_VAR
VAR CONSTANT
    DL_STEP_MAX  : INT := 32;                      // 步骤数上限 [步] / Step count limit
    DL_STEP_MIN  : INT := 1;                       // 步骤数下限 [步] / Step count lower bound
    DL_SEC_MS    : TIME := T#1S;                   // 一秒基准 [毫秒] / One second base
    DL_TIME_ZERO : TIME := T#0S;                   // 时间零值基准 [毫秒] / Time zero reference
    DL_TIME_MIN  : TIME := T#1MS;                  // 时间参数最小正值 [毫秒] / Minimum positive time
END_VAR

(*------------------------------------------------------------------------------
 * 段 1｜输出确定性默认值（单拍标志每拍预清零，R25 第一律）
 *      Deterministic defaults first, one-scan flags pre-cleared every scan
 *-----------------------------------------------------------------------------*)
bRequestStep  := FALSE;                         // 步骤请求单拍预清零（Step request pulse pre-cleared）
bRequestAbort := FALSE;                         // 中止请求单拍预清零（Abort request pulse pre-cleared）
uInfoCode     := 16#0000_0000;                  // 信息级码每拍重算（Info code recomputed every scan）
bCmdDropped   := FALSE;                         // 丢弃标记预清零（Dropped flag pre-cleared）
bSecTick      := FALSE;                         // 秒脉冲预清零（Second tick pre-cleared）

(*------------------------------------------------------------------------------
 * 段 2｜沿检测无条件刷新（红线：实例在 CASE 之外每拍必刷）
 *      Edge detection refreshed unconditionally outside the CASE
 *-----------------------------------------------------------------------------*)
fbTrigStart(CLK := bStart);
fbTrigHold(CLK := bHold);
fbTrigRestart(CLK := bRestart);
fbTrigStop(CLK := bStop);
fbTrigAbort(CLK := bAbort);
fbTrigReset(CLK := bReset);
fbTrigStepDone(CLK := bStepDone);

(*------------------------------------------------------------------------------
 * 段 3｜首扫初始化（唯一合法范式：初值 FALSE，判据取非）
 *      First-scan initialisation following the single legal pattern
 *-----------------------------------------------------------------------------*)
IF NOT bInit THEN
    nStep         := 0;                         // 步骤号清零（Step number cleared）
    nStepUse      := DL_STEP_MIN;               // 生效步骤数取下限（Effective step count at the lower bound）
    bStepIssued   := FALSE;                     // 请求已发出标志清零（Request issued flag cleared）
    bStepAcked    := FALSE;                     // 完成已消费标志清零（Completion consumed flag cleared）
    bHoldArmed    := FALSE;                     // 暂停登记清零（Hold armed cleared）
    bStopArmed    := FALSE;                     // 停止登记清零（Stop armed cleared）
    uElapsed      := 0;                         // 运行秒累计清零（Elapsed seconds cleared）
    bFaultLatch   := FALSE;                     // 故障锁存清零（Fault latch cleared）
    uErrInt       := 16#0000_0000;              // 故障码清零（Fault code cleared）
    eState        := E_DL_BatchPhaseState.eIdle; // 相状态复位为空闲（Phase state reset to idle）
    ePhase        := E_DL_BatchPhaseState.eIdle; // 状态出口复位（State outlet reset）
    nStepNo       := 0;                         // 步骤号出口清零（Step outlet cleared）
    uPhaseElapsed := 0;                         // 累计时间出口清零（Elapsed outlet cleared）
    bError        := FALSE;                     // 故障位出口清零（Fault outlet cleared）
    bInit         := TRUE;                      // 首扫只做一次（First scan runs once）
END_IF

(*------------------------------------------------------------------------------
 * 段 4｜参数钳位（步骤数越界属组态，钳位加信息码，不停机）
 *      Parameter clamping with an informational code only
 *-----------------------------------------------------------------------------*)
IF nStepCount < DL_STEP_MIN THEN
    nStepUse  := DL_STEP_MIN;                   // 步骤数下限钳位（Clamped to the lower bound）
    uInfoCode := 16#0005_0104;                  // 0104 步骤数越界已钳位（Step count clamped）
ELSIF nStepCount > DL_STEP_MAX THEN
    nStepUse  := DL_STEP_MAX;                   // 步骤数上限钳位（Clamped to the upper bound）
    uInfoCode := 16#0005_0104;                  // 0104 步骤数越界已钳位（Step count clamped）
ELSE
    nStepUse  := nStepCount;                    // 合法步骤数直通（Valid step count passed through）
END_IF

IF tStepTimeout <= DL_TIME_ZERO THEN
    tStepUse  := DL_TIME_MIN;                   // 零表示关闭监控，定时器仍给安全预置值（Zero disables, the timer keeps a safe preset）
    bStepMon  := FALSE;                         // 单步监控关闭（Step watchdog disabled）
    uInfoCode := 16#0005_0107;                  // 0107 单步超时监控关闭（Step watchdog disabled）
ELSE
    tStepUse  := tStepTimeout;                  // 合法超时直通（Valid timeout passed through）
    bStepMon  := TRUE;                          // 单步监控启用（Step watchdog enabled）
END_IF

IF tHoldTimeout <= DL_TIME_ZERO THEN
    tHoldUse  := DL_TIME_MIN;                   // 零表示关闭监控（Zero disables the watchdog）
    bHoldMon  := FALSE;                         // 暂停监控关闭（Hold watchdog disabled）
    uInfoCode := 16#0005_0107;                  // 0107 暂停超时监控关闭（Hold watchdog disabled）
ELSE
    tHoldUse  := tHoldTimeout;                  // 合法超时直通（Valid timeout passed through）
    bHoldMon  := TRUE;                          // 暂停监控启用（Hold watchdog enabled）
END_IF
IF nStep < 0 THEN
    nStep := 0;                                 // 步骤号负值防御，正常流程不可达（Defensive clamp, unreachable normally）
END_IF

(*------------------------------------------------------------------------------
 * 段 5｜命令优先级裁决（中止 高于 停止 高于 暂停 高于 恢复 高于 启动；不排队）
 *      Command arbitration by a strict priority order, dropped commands are not queued
 *-----------------------------------------------------------------------------*)
bCmdAbort   := fbTrigAbort.Q;                   // 最高优先：中止（Highest priority, abort）
bCmdStop    := fbTrigStop.Q AND (NOT bCmdAbort); // 次优先：停止（Next, stop）
bCmdHold    := fbTrigHold.Q AND (NOT bCmdAbort) AND (NOT bCmdStop); // 次优先：暂停（Next, hold）
bCmdRestart := fbTrigRestart.Q AND (NOT bCmdAbort) AND (NOT bCmdStop) AND (NOT bCmdHold); // 次优先：恢复（Next, restart）
bCmdStart   := fbTrigStart.Q AND (NOT bCmdAbort) AND (NOT bCmdStop) AND (NOT bCmdHold) AND (NOT bCmdRestart); // 最低优先：启动（Lowest, start）
bCmdReset   := fbTrigReset.Q;                   // 复位独立通道，不参与优先级（Reset is an independent channel）

IF (bCmdAbort AND (fbTrigStop.Q OR fbTrigHold.Q OR fbTrigRestart.Q OR fbTrigStart.Q)) OR
   (bCmdStop AND (fbTrigHold.Q OR fbTrigRestart.Q OR fbTrigStart.Q)) OR
   (bCmdHold AND (fbTrigRestart.Q OR fbTrigStart.Q)) OR
   (bCmdRestart AND fbTrigStart.Q) THEN
    bCmdDropped := TRUE;                        // 同拍多命令：标记丢弃提示（Concurrent commands, mark the drop）
END_IF
IF bCmdDropped THEN
    uInfoCode := 16#0005_0105;                  // 0105 低优先命令已丢弃（Low priority command dropped）
END_IF

(*------------------------------------------------------------------------------
 * 段 6｜定时器无条件刷新（入口条件取当前相状态；掉使能时冻结计时）
 *      Timers refreshed unconditionally, gated by enable and by the phase state
 *-----------------------------------------------------------------------------*)
fbStepWatch(IN := bEnable AND bStepMon AND (NOT bStepWatchBreak) AND
                 ((eState = E_DL_BatchPhaseState.eRunning) OR
                  (eState = E_DL_BatchPhaseState.eCompleting) OR
                  (eState = E_DL_BatchPhaseState.eStopping)),
            PT := tStepUse);
bStepTo := fbStepWatch.Q;                       // 超时判定在实例调用后取用（Verdict read after the call）
bStepWatchBreak := FALSE;                       // 断输入脉冲在实例调用后自清（Break pulse self-cleared after the call）

fbHoldWatch(IN := bEnable AND bHoldMon AND (eState = E_DL_BatchPhaseState.eHeld), PT := tHoldUse);
bHoldTo := fbHoldWatch.Q;                       // 超时判定在实例调用后取用（Verdict read after the call）

fbSecBase(IN := bEnable AND (NOT bSecDone), PT := DL_SEC_MS);
bSecTick := fbSecBase.Q;                        // 秒脉冲在实例调用后取用（Tick read after the call）
bSecDone := fbSecBase.Q;                        // 到点电平在实例调用后更新，供下拍自复位（Elapsed level refreshed after the call）

(*------------------------------------------------------------------------------
 * 段 7｜主状态机（枚举每个成员均有标签，末尾 ELSE 兜底到已中止）
 *      Main state machine, one label per member plus a trailing ELSE fallback
 *      掉使能时整体冻结：状态、步骤号与单拍请求都不变（A disabled phase is frozen）
 *-----------------------------------------------------------------------------*)
IF bEnable THEN
    CASE eState OF

        E_DL_BatchPhaseState.eIdle: // 空闲：等启动，输出全复位
            nStep        := 0;              // 步骤号归零（Step number cleared）
            bStepIssued  := FALSE;          // 请求标志清零（Request flag cleared）
            bStepAcked   := FALSE;          // 完成消费标志清零（Completion flag cleared）
            bHoldArmed   := FALSE;          // 暂停登记清零（Hold armed cleared）
            bStopArmed   := FALSE;          // 停止登记清零（Stop armed cleared）
            IF bCmdStart THEN
                nStep       := 1;           // 从第一步开始（Start from the first step）
                bStepIssued := FALSE;       // 请求待下拍发出（The request is issued on the next scan）
                eState      := E_DL_BatchPhaseState.eRunning; // 进执行相（Enter the running phase）
            END_IF

        E_DL_BatchPhaseState.eRunning: // 执行：推进步骤，处理四类命令
            IF bCmdAbort THEN
                bHoldArmed := FALSE;        // 中止优先：清暂停登记（Abort wins, clear the hold armed flag）
                bStopArmed := FALSE;        // 清停止登记（Clear the stop armed flag）
                eState     := E_DL_BatchPhaseState.eAborting; // 进中止相（Enter the aborting phase）
            ELSIF bStepFail THEN
                IF NOT bFaultLatch THEN
                    bFaultLatch := TRUE;    // 步骤失败：锁故障（Step failure, latch the fault）
                    uErrInt     := 16#0005_0204; // 0204 步骤失败（Step failure）
                END_IF
                eState := E_DL_BatchPhaseState.eAborting; // 进中止相（Enter the aborting phase）
            ELSIF bCmdHold THEN
                bHoldArmed := TRUE;         // 受理暂停，寄存器置位（The hold request is accepted）
                IF NOT bStepIssued THEN
                    eState := E_DL_BatchPhaseState.eHeld;    // 本步尚未开始：直接暂停（The step has not started, hold at once）
                ELSE
                    eState := E_DL_BatchPhaseState.eHolding; // 本步进行中：等步骤边界（Wait for the step boundary）
                END_IF
            ELSE
                IF bCmdStop THEN
                    bStopArmed := TRUE;     // 登记停止，在步骤边界生效（Arm the stop at the boundary）
                END_IF
                IF fbTrigStepDone.Q AND (NOT bStepAcked) THEN
                    bStepAcked  := TRUE;    // 消费本次完成（Consume the completion）
                    bStepIssued := FALSE;   // 下一步的请求待重新发出（The next step needs a new request）
                    bStepWatchBreak := TRUE; // 步骤边界：单步超时断输入一拍，按步重计时（Restart the step watchdog at the boundary）
                    IF bStopArmed THEN
                        eState := E_DL_BatchPhaseState.eStopping; // 边界已到：进停止相（Boundary reached, stop）
                    ELSIF nStep >= nStepUse THEN
                        eState := E_DL_BatchPhaseState.eCompleting; // 步骤耗尽：进收尾相（Steps exhausted, complete）
                    ELSE
                        nStep := nStep + 1; // 推进到下一步（Advance to the next step）
                    END_IF
                ELSIF bStepTo THEN
                    IF NOT bFaultLatch THEN
                        bFaultLatch := TRUE; // 单步超时：锁故障（Step timeout, latch the fault）
                        uErrInt     := 16#0005_0203; // 0203 单步超时（Step timeout）
                    END_IF
                    eState := E_DL_BatchPhaseState.eAborting; // 进中止相（Enter the aborting phase）
                ELSE
                    IF bStepDone THEN
                        bStepAcked := TRUE;  // 反馈仍高：保持已消费（Feedback still high, keep the consumed flag）
                    ELSE
                        bStepAcked := FALSE; // 反馈落下：允许下一次消费（Feedback dropped, allow the next consumption）
                    END_IF
                    IF NOT bStepIssued THEN
                        bRequestStep := TRUE; // 单拍步骤请求（One-scan step request）
                        bStepIssued  := TRUE; // 置请求已发（Mark the request as issued）
                    END_IF
                END_IF
            END_IF

        E_DL_BatchPhaseState.eCompleting: // 收尾：等收尾动作反馈，不占步骤号
            IF bCmdAbort THEN
                eState := E_DL_BatchPhaseState.eAborting; // 中止优先（Abort wins）
            ELSIF bStepFail THEN
                IF NOT bFaultLatch THEN
                    bFaultLatch := TRUE;    // 收尾失败：锁故障（Clean-up failure, latch the fault）
                    uErrInt     := 16#0005_0204; // 0204 步骤失败（Step failure）
                END_IF
                eState := E_DL_BatchPhaseState.eAborting; // 进中止相（Enter the aborting phase）
            ELSIF fbTrigStepDone.Q AND (NOT bStepAcked) THEN
                bStepAcked := TRUE;         // 收尾完成（Clean-up finished）
                eState     := E_DL_BatchPhaseState.eComplete; // 进完成相（Enter the complete phase）
            ELSIF bStepTo THEN
                IF NOT bFaultLatch THEN
                    bFaultLatch := TRUE;    // 收尾超时：锁故障（Clean-up timeout, latch the fault）
                    uErrInt     := 16#0005_0203; // 0203 单步超时（Step timeout）
                END_IF
                eState := E_DL_BatchPhaseState.eAborting; // 进中止相（Enter the aborting phase）
            ELSE
                IF bStepDone THEN
                    bStepAcked := TRUE;     // 反馈仍高：保持已消费（Feedback still high）
                ELSE
                    bStepAcked := FALSE;    // 反馈落下：允许下一次消费（Feedback dropped）
                END_IF
            END_IF

        E_DL_BatchPhaseState.eComplete: // 完成：保持到复位，已终止态不受理启动与中止
            bStepIssued := FALSE;           // 终止态不保留步骤请求标志（No step request lingers in a terminal state）

        E_DL_BatchPhaseState.eHolding: // 暂停请求：仅在步骤边界真正暂停
            IF bCmdAbort THEN
                eState := E_DL_BatchPhaseState.eAborting; // 中止优先（Abort wins）
            ELSIF bCmdStop THEN
                bStopArmed := TRUE;         // 停止优先于暂停（Stop outranks hold）
                eState     := E_DL_BatchPhaseState.eStopping; // 进停止相（Enter the stopping phase）
            ELSIF bHoldArmed AND (NOT bStepIssued) THEN
                eState := E_DL_BatchPhaseState.eHeld; // 步骤尚未开始：可安全暂停（The step has not started, safe to hold）
            ELSIF fbTrigStepDone.Q AND (NOT bStepAcked) THEN
                bStepAcked  := TRUE;        // 当前步完成反馈到达：边界已到（The boundary has arrived）
                bStepIssued := FALSE;       // 清请求标志（Clear the issued flag）
                eState      := E_DL_BatchPhaseState.eHeld; // 进已暂停相（Enter the held phase）
            ELSE
                IF bStepDone THEN
                    bStepAcked := TRUE;     // 反馈仍高：保持已消费（Feedback still high）
                ELSE
                    bStepAcked := FALSE;    // 反馈落下：允许下一次消费（Feedback dropped）
                END_IF
            END_IF

        E_DL_BatchPhaseState.eHeld: // 已暂停：不推进、不发请求
            IF bCmdAbort THEN
                eState := E_DL_BatchPhaseState.eAborting; // 中止优先（Abort wins）
            ELSIF bCmdStop THEN
                bStopArmed := TRUE;         // 登记停止（Arm the stop）
                eState     := E_DL_BatchPhaseState.eStopping; // 进停止相（Enter the stopping phase）
            ELSIF bCmdRestart THEN
                bStepIssued := FALSE;       // 恢复：请求待重发（Restart, the request is reissued）
                bStepAcked  := FALSE;       // 恢复：重新等待本步完成反馈（Restart, wait for a fresh completion）
                eState      := E_DL_BatchPhaseState.eRestarting; // 进恢复相（Enter the restarting phase）
            ELSIF bHoldTo THEN
                IF NOT bFaultLatch THEN
                    bFaultLatch := TRUE;    // 暂停超时：锁故障（Hold timeout, latch the fault）
                    uErrInt     := 16#0005_0205; // 0205 暂停超时（Hold timeout）
                END_IF
                eState := E_DL_BatchPhaseState.eAborting; // 进中止相（Enter the aborting phase）
            ELSE
                bHoldArmed := TRUE;         // 保持登记，等待恢复或停止（Keep the hold armed）
            END_IF

        E_DL_BatchPhaseState.eRestarting: // 恢复中：重发当前步请求，不重头
            bRequestStep := TRUE;           // 重发当前步请求（Reissue the current step request）
            bStepIssued  := TRUE;           // 置请求已发（Mark the request as issued）
            bStepAcked   := FALSE;          // 重新等待本步完成（Wait for a fresh completion）
            uInfoCode    := 16#0005_0106;   // 0106 从暂停恢复，步骤号不重置（Restarted from hold, the step number is kept）
            eState       := E_DL_BatchPhaseState.eRunning; // 回执行相（Back to running）

        E_DL_BatchPhaseState.eStopping: // 停止中：等收尾反馈
            IF bCmdAbort THEN
                eState := E_DL_BatchPhaseState.eAborting; // 中止优先（Abort wins）
            ELSIF fbTrigStepDone.Q AND (NOT bStepAcked) THEN
                bStepAcked := TRUE;         // 收尾完成（Wrap-up finished）
                eState     := E_DL_BatchPhaseState.eStopped; // 进已停相（Enter the stopped phase）
            ELSIF bStepTo THEN
                IF NOT bFaultLatch THEN
                    bFaultLatch := TRUE;    // 收尾超时：锁故障（Wrap-up timeout, latch the fault）
                    uErrInt     := 16#0005_0203; // 0203 单步超时（Step timeout）
                END_IF
                eState := E_DL_BatchPhaseState.eAborting; // 进中止相（Enter the aborting phase）
            ELSE
                IF bStepDone THEN
                    bStepAcked := TRUE;     // 反馈仍高：保持已消费（Feedback still high）
                ELSE
                    bStepAcked := FALSE;    // 反馈落下：允许下一次消费（Feedback dropped）
                END_IF
            END_IF

        E_DL_BatchPhaseState.eStopped: // 已停：保持到复位，已终止态不受理启动与中止
            bStepIssued := FALSE;           // 终止态不保留步骤请求标志（No step request lingers in a terminal state）

        E_DL_BatchPhaseState.eAborting: // 中止中：发出中止动作单拍后立即进已中止
            bRequestAbort := TRUE;          // 单拍中止动作请求（One-scan abort action request）
            bHoldArmed    := FALSE;         // 清暂停登记（Clear the hold armed flag）
            bStopArmed    := FALSE;         // 清停止登记（Clear the stop armed flag）
            eState        := E_DL_BatchPhaseState.eAborted; // 进已中止相（Enter the aborted phase）

        E_DL_BatchPhaseState.eAborted: // 已中止：保持到复位，步骤号保留供报表追溯
            bStepIssued := FALSE;           // 终止态不保留步骤请求标志（No step request lingers in a terminal state）

        ELSE
            bFaultLatch := TRUE;            // 非法状态兜底锁存（Illegal state latched）
            uErrInt     := 16#0005_0206;    // 0206 非法状态兜底（Illegal state fallback code）
            eState      := E_DL_BatchPhaseState.eAborted; // 直接进已中止，不回空闲（Go straight to aborted）
    END_CASE

    (* 秒脉冲累加：只在执行相计时，暂停与收尾不计入相净运行时间 *)
    IF bSecTick AND (eState = E_DL_BatchPhaseState.eRunning) THEN
        uElapsed := uElapsed + 1;           // 相净运行秒累加（Accumulate a running second）
    END_IF
END_IF

(*------------------------------------------------------------------------------
 * 段 8｜复位（仅已终止态受理；清步骤号、完成标志与故障锁存）
 *      Reset is accepted from the terminal states only
 *-----------------------------------------------------------------------------*)
IF bCmdReset THEN
    IF (eState = E_DL_BatchPhaseState.eComplete) OR (eState = E_DL_BatchPhaseState.eStopped) OR
       (eState = E_DL_BatchPhaseState.eAborted) OR (eState = E_DL_BatchPhaseState.eIdle) THEN
        nStep       := 0;                   // 步骤号归零（Step number cleared）
        bStepIssued := FALSE;               // 请求标志清零（Request flag cleared）
        bStepAcked  := FALSE;               // 完成消费标志清零（Completion flag cleared）
        bHoldArmed  := FALSE;               // 暂停登记清零（Hold armed cleared）
        bStopArmed  := FALSE;               // 停止登记清零（Stop armed cleared）
        bFaultLatch := FALSE;               // 清故障锁存（Clear the fault latch）
        uErrInt     := 16#0000_0000;        // 清故障码（Clear the fault code）
        eState      := E_DL_BatchPhaseState.eIdle; // 回空闲（Back to idle）
    END_IF
END_IF

(*------------------------------------------------------------------------------
 * 段 9｜出口映射（状态、步骤号、活动族、完成标志、累计时间与码位定级）
 *      Outlet mapping with a single priority chain for the event code
 *-----------------------------------------------------------------------------*)
ePhase        := eState;                        // 相状态出口（Phase state outlet）
nStepNo       := nStep;                         // 步骤号出口（Step number outlet）
uPhaseElapsed := uElapsed;                      // 净运行时间出口（Elapsed outlet）
bPhaseComplete := (eState = E_DL_BatchPhaseState.eComplete); // 完成标志由状态派生（Derived from the state）
bPhaseActive  := (eState = E_DL_BatchPhaseState.eRunning) OR
                 (eState = E_DL_BatchPhaseState.eCompleting) OR
                 (eState = E_DL_BatchPhaseState.eHolding) OR
                 (eState = E_DL_BatchPhaseState.eHeld) OR
                 (eState = E_DL_BatchPhaseState.eRestarting) OR
                 (eState = E_DL_BatchPhaseState.eStopping) OR
                 (eState = E_DL_BatchPhaseState.eAborting); // 活动族派生（Active family derived）
bError        := bFaultLatch;                   // 故障位只反映故障级锁存（Fault bit reflects the latch only）
IF bError THEN
    uErrorId := uErrInt;                        // 故障级码优先透出（Fault level code has priority）
ELSE
    uErrorId := uInfoCode;                      // 无故障透出本拍信息级码（Info code exposed otherwise）
END_IF
END_FUNCTION_BLOCK

(* ---- FB_DL_BatchTransferSeq.st ---- *)
(*==============================================================================
 * 组件名称 (Component)  : FB_DL_BatchTransferSeq
 * 溯源说明 (Provenance): 道莅 clean-room 防御性实现（IEC 61131-3 纯净实现，闭源文档仅借语义，零代码行）
 * 所属子库 (Sublibrary) : DL_Process / Sequence
 * 当前版本 (Version)    : 1.0.2
 * 兼容性   (Platform)   : CODESYS 3.5 / TwinCAT 3 / 汇川 InoProShop / 施耐德
 *                         Machine Expert；纯 IEC 61131-3（第 3 版），仅用
 *                         Standard.library 的 TON / TIME_TO_DINT / DINT_TO_TIME
 * 组件分类 (Category)   : 功能块（FUNCTION_BLOCK）· 批次物料转移顺控
 * 功能一句话 (Summary)  : 开阀 → 等双阀开到位 → 启泵 → 计量转移 → 停泵 →
 *                         排空验证 → 关阀，按 ISA-88 相/步骤最小语义编排。
 *
 * 本件存在的意义 (Why this unit exists)
 *   批次转移是 ISA-88 相步骤的最小实证单元，也是 OEE 事故的高发点：
 *   泵在阀没到位时就启（干转烧泵）、中止时先关阀后停泵（管道憋压）、
 *   转移量靠程序自己积分（累计量双份口径，对不上账）。本件把这三件事
 *   写成结构约束：泵的启动条件是双阀反馈、中止路径先停泵再关阀、
 *   累计量**由调用方积分器注入**，本件不重复积分。
 *
 * 步骤与判据 (Steps and criteria)
 *   ePrepValve   : 双阀开指令，等 bSrcValveFb 与 bDstValveFb **同时**到位
 *   eTransferring: 双阀保持、泵启动；fTransferred >= fVolumeTarget → 停泵
 *   eDraining    : 泵停、双阀仍开；fFlow < fDrainFlow 持续 tDrainVerify → 判排空完成
 *   eClosing     : 双阀关指令（本库阀门指令语义：TRUE = 开启，故关阀 = 清指令），
 *                  等关阀确认窗（tValveFb）后进 eComplete
 *   eComplete    : 放行；bStart 落下才回 eIdle（不自动开始下一批）
 *   eAbort       : 中止兼容路径（xCoastStop = FALSE）：先停泵后关阀（顺序
 *                  不可反，防管道憋压），等 bStart 落下复位
 *   eAbortCoast  : 中止第一段（xCoastStop = TRUE，推荐）：泵输出使能立即断、
 *                  **阀位保持不动**（不发关阀指令），泵惰转计时窗内管路
 *                  残压随泵惰转泄放，杜绝停泵与关阀同拍发出的物理竞态
 *   eAbortClose  : 中止第二段：惰转窗满后发关阀指令（清阀门指令），等阀
 *                  离开开位（双阀开反馈任一保持即计时）；确认超时 → 0317
 *
 * 中止语义（三件顺控件共用同一段口径）
 *   bAbort **任意拍**生效（中止族态内不重复触发，防惰转窗被反复重启）：
 *   xCoastStop = TRUE 走两段化——段 A 断泵输出使能、阀保持不动、惰转计时；
 *   段 B 惰转窗满发关阀指令，等关阀确认，超时报 0317。两段之间由 TON 跨拍
 *   物理时序分隔，**禁止单拍内「停泵赋值 + 关阀赋值」连续成立**（机检断言：
 *   abort 拍不得出现关阀输出置位）。xCoastStop = FALSE 保留 v1.0.1 单拍
 *   行为（仅存量调用兼容，**不推荐：泵惰转期间残压可经未关阀位回流**）。
 *   中止**不排队、不回退重来、不自动续跑**——中止是人的决定，重启必须由
 *   新的 bStart 重新开始。bStart 落沿同样按中止处理（外部撤销）。
 *
 * 边界安全 (Boundary)
 *   ① fVolumeTarget <= 0 或 tTimeout = T#0S → 故障 0315、停泵关阀、回 eFault；
 *   ② 阀位反馈超 tValveFb 未到位 → 故障 0314、**不启泵**、回 eIdle 并先清输出；
 *   ③ 转移总时长超 tTimeout → 故障 0315（复用，R90）；
 *   ④ fTransferred 由调用方注入：**批次切换必须由调用方清零累计器**；本件以本拍
 *      值为准，不做回退检测（回退是换批的正常现象，不是故障，若在此报错会
 *      让每批首拍都报一次假故障）；该口径以信息 01E0 在进入转移相时声明一次；
 *   ⑤ 输入非有限（累计量或流量）→ 复用 0315 并停泵关阀（无专用码位，R90）；
 *   ⑥ 泵/阀三输出互斥在段 1 全清、段 7 按相置位（R72 双路径）；
 *   ⑦ 四只 TON 各司其职：开阀到位 / 关阀确认 / 排空验证 / 总时长，
 *      绝不复用同一实例跨相计时（R40；规格写三个实例，关阀确认必须独立，故实测为四只）；
 *      v1.0.2 增至六只：惰转计时 / 中止关阀确认各自独立实例，同样不复用；
 *   ⑧ CASE 落 ELSE 置 0316 并回 eFault；
 *   ⑨ xCoastStop = TRUE 且 tPumpCoastTime <= 0 → 参数非法 0315 复用（R90：
 *      惰转窗为 0 使两段化退化为单拍，违背修复意图，按非法参数拦截）。
 *
 * 验收向量（v1.0.2 中止时序，修复后必测）：
 *   V9  abort 触发拍（xCoastStop = TRUE）：泵指令 FALSE、双阀指令保持开
 *       （TRUE）、关阀输出（指令清零动作）当拍不发生——机检断言主向量；
 *   V10 惰转窗未满期间跨拍扫描：双阀指令恒保持开、泵指令恒 FALSE
 *       （跨拍验证，窗内无任何输出翻转）；
 *   V11 惰转窗满拍：双阀指令置 FALSE（发关阀指令）；
 *   V12 关阀确认超时（阀开反馈在确认窗内仍保持）→ eErr = 16#0005_0317
 *       且 bError 置位（R45 配对），输出保持关阀指令；
 *   V13 xCoastStop = FALSE：回归 v1.0.1 向量 V4（abort 拍泵 FALSE 且阀
 *       指令 FALSE 同拍成立，兼容路径单拍中止）。
 *
 * 错误码    : 16#0005_01E0 累计转移量由调用方积分器注入，本件不重复积分——信息级，口径声明
 *             16#0005_01E1 排空验证窗内流量持续低于门限，判排空完成——信息级，正常结论
 *             16#0005_0314 阀位反馈超时未到位，拒绝启泵——故障级，回 eIdle 并先清输出
 *             16#0005_0315 转移总时长超时或体积/超时/输入参数非法（含非有限复用，R90）——故障级
 *             16#0005_0316 状态机落 ELSE 兜底（非法状态）——故障级，回 eFault 并先清输出
 *             16#0005_0317 中止第二段关阀确认超时（阀开反馈在确认窗内保持，
 *                          v1.0.2 新增）——故障级，置 bError，保持关阀指令等启动撤销
 * 码位总账  : 16#0005_01E0 用 / 16#0005_01E1 用 ｜ 16#0005_0314 用 / 16#0005_0315 用 /
 *             16#0005_0316 用 / 16#0005_0317 用（R23 特批故障槽）
 * 状态机    : E_DL_TransferState（eIdle / ePrepValve / eTransferring / eDraining / eClosing /
 *             eComplete / eAbort / eAbortCoast / eAbortClose / eFault），
 *             CASE 含 ELSE 兜底，ELSE 置 16#0005_0316 并回 eFault
 * 采样约定  : 每任务周期调用一次；各窗时长由引脚给定，不读系统时钟
 * 依赖说明  : 只做组合编排；累计量由调用方以 FB_DL_Integrator 注入，本件**不内联积分**
 * 验收向量  : V1 双阀反馈到位 → 泵启动（启泵条件主向量）；fTransferred 达 5.0 m³ → 停泵
 *             V2 阀位反馈 5 s 内未到位 → 0314，泵始终 FALSE，回 eIdle（不启泵主向量）
 *             V3 排空相流量 0.02 m³/h（< 0.05）持续 10 s → bDrained = TRUE，eErr = 01E1 → eClosing
 *             V4 转移中 bAbort → 同拍泵 FALSE 且阀指令 FALSE，回 eAbort（中止主向量）
 *             V5 转移总时长超 30 min → 0315，停泵关阀，bFailed = TRUE
 *             V6 fVolumeTarget = 0 → 0315，回 eFault，bValid = FALSE
 *             V7 fTransferred = NaN → 0315 复用，停泵关阀（坏值安全侧）
 *             V8 换批（fTransferred 由 5.0 回 0.1）→ **不报故障**，以本拍值为准继续（口径主向量）
 * 红线自检  : 全局变量声明零使用 / 外部变量访问零使用 / 物理地址零使用 ｜ 纯 IEC 61131-3 ｜ 无除法
 *             浮点只用大小比较 ｜ 无循环 ｜ 全变量双语同行注释 ｜ ENUM + CASE 含 ELSE
 *             ｜ 六只 TON 在主体前部无条件刷新 ｜ 单拍标志全部预清零 ｜ 阈值常量化
 * 修订历史  : 2026-11-16  v1.0.0  首版入库（R22 · 批 3 · 批处理顺控）
 *             2026-11-16  v1.0.1  R22 终审修复：总时长超时分支（0315）补置
 *             bError := TRUE——故障级码位必须同时置故障标志（R45 纪律），
 *             原实现只给码不置标志，bValid 误判为可用
 *             2026-11-17  v1.0.2  R23 P0 修复：中止时序两段化——新增
 *             xCoastStop（默认 TRUE 走惰转两段化）与 tPumpCoastTime（惰转
 *             窗）引脚；段 A 断泵输出使能、阀位保持不动、惰转计时；段 B
 *             窗满发关阀指令、确认超时置新故障码 16#0005_0317 + bError
 *             （R45 配对）；禁止单拍「停泵 + 关阀」连续成立；验收向量
 *             V9~V13 收录于本头注释「验收向量（v1.0.2 中止时序）」段；xCoastStop = FALSE 保留 v1.0.1
 *             单拍行为（不推荐：残压回流风险）
 *============================================================================*)

(*-----------------------------------------------------------------------------
 * 枚举: E_DL_TransferState（归属本功能块，同文件发布，全库唯一定义）
 * 含义: 批次转移顺控相位，每个成员在 CASE 中有且仅有一个标签。
 *-----------------------------------------------------------------------------*)
TYPE E_DL_TransferState :
(
    eIdle         := 0,   // 待机：未启动 / Idle, not started
    ePrepValve    := 10,  // 准备阀门：双阀开指令，等开到位反馈 / Preparing, valves open, waiting for feedback
    eTransferring := 20,  // 转移中：泵运行，按注入累计量判结束 / Transferring, the pump runs
    eDraining     := 30,  // 排空中：泵停，等流量降到门限以下 / Draining, the pump stopped
    eClosing      := 40,  // 关阀中：双阀关指令，等确认窗 / Closing, waiting for the confirmation window
    eComplete     := 50,  // 完成：放行 / Complete, released
    eAbort        := 60,  // 中止兼容路径：单拍停泵关阀（xCoastStop = FALSE，不推荐） / Legacy single-scan abort, pump and valves off in one scan
    eAbortCoast   := 61,  // 中止第一段：泵输出使能已断，阀位保持不动，惰转计时中 / Abort stage A, pump disabled, valves held, coast timing
    eAbortClose   := 62,  // 中止第二段：惰转窗满，关阀指令已发，等阀离开开位 / Abort stage B, close command issued, waiting for the valve to leave open position
    eFault        := 99   // 故障：参数/超时/非法状态 / Fault, parameters, timeout or an illegal state
);
END_TYPE

FUNCTION_BLOCK FB_DL_BatchTransferSeq
VAR_INPUT
    bStart        : BOOL;                      // 启动请求，电平有效 / start request, level active
    bAbort        : BOOL;                      // 中止请求，任意拍生效 / abort request, effective on any scan
    bSrcValveFb   : BOOL;                      // 源阀开到位反馈 / source valve open feedback
    bDstValveFb   : BOOL;                      // 目标阀开到位反馈 / destination valve open feedback
    fTransferred  : REAL;                      // 累计转移量 [m3]，**由调用方积分器注入** / transferred volume, injected by the caller
    fVolumeTarget : REAL := 5.0;               // 目标转移量 [m3]，须 > 0 / target volume [m3], must be > 0
    fFlow         : REAL;                      // 实测流量 [m3/h] / measured flow [m3/h]
    fDrainFlow    : REAL := 0.05;              // 排空判据流量门限 [m3/h] / drain flow threshold [m3/h]
    tDrainVerify  : TIME := T#10S;             // 排空验证时长 [ms] / drain verification duration [ms]
    tValveFb      : TIME := T#5S;              // 阀位反馈确认窗 [ms] / valve feedback window [ms]
    tTimeout      : TIME := T#30M;             // 转移总时长上限 [ms]，须 > 0 / total transfer timeout [ms], must be > 0
    xCoastStop    : BOOL := TRUE;              // TRUE = 中止走惰转两段化（推荐）/ FALSE = 兼容旧行为单拍中止（仅存量调用保留，不推荐：残压回流风险） / Coast-stop abort sequencing enabled
    tPumpCoastTime: TIME := T#2S;              // 泵惰转时间 [ms]（默认 2 s）：停泵到关阀的物理时序分隔窗 / Pump coast-down time [ms]
END_VAR
VAR_OUTPUT
    bPumpCmd      : BOOL;                      // 泵指令 / pump command
    bSrcValveCmd  : BOOL;                      // 源阀指令（TRUE = 开启） / source valve command, TRUE means open
    bDstValveCmd  : BOOL;                      // 目标阀指令（TRUE = 开启） / destination valve command
    bDrained      : BOOL;                      // 排空完成标志 / drained flag
    bDone         : BOOL;                      // 转移完成放行 / transfer complete, released
    bFailed       : BOOL;                      // 转移失败锁定 / transfer failed, latched
    eErr          : UDINT;                     // 错误码，0 表示无错 / error code, 0 means no error
    bError        : BOOL;                      // 故障级标志，仅故障级错误置位 / fault-class flag, set only on fault-level codes
    bValid        : BOOL;                      // 输出可用标志 / outputs usable flag
END_VAR
VAR
    fbValveFb     : TON;                       // 开阀到位确认窗，段 6 无条件刷新 [ms] / open feedback window
    fbCloseFb     : TON;                       // 关阀确认窗，段 6 无条件刷新 [ms] / close confirmation window
    fbDrain       : TON;                       // 排空验证窗，段 6 无条件刷新 [ms] / drain verification window
    fbTotal       : TON;                       // 转移总时长，段 6 无条件刷新 [ms] / total transfer timer
    fbCoast       : TON;                       // 泵惰转计时窗（中止第一段），段 6 无条件刷新 [ms] / pump coast-down window, abort stage A
    fbAbortClose  : TON;                       // 中止关阀确认窗（中止第二段，独立实例不复用），段 6 无条件刷新 [ms] / abort close-confirm window, stage B, dedicated instance
    _eState       : E_DL_TransferState := E_DL_TransferState.eIdle; // 当前相位 / current phase
    _bInit        : BOOL := FALSE;             // 首扫标志，初值 FALSE 取非判定 / first-scan flag, tested negated
    _bParamBad    : BOOL;                      // 参数非法标志 / illegal parameter flag
    _bFiniteBad   : BOOL;                      // 输入非有限标志 / non-finite input flag
    _bIllegal     : BOOL;                      // 非法状态标志 / illegal state flag
    _bFaultAcc    : BOOL;                      // 故障锁存保持量（等新启动清除） / held fault latch, cleared by a new start
    _bFailedAcc   : BOOL;                      // 失败锁存保持量 / held failure latch
    _bBothFb      : BOOL;                      // 双阀同时到位 / both valves reported open
    _bDrainCond   : BOOL;                      // 排空条件（流量低于门限） / drain condition
    _bFbBreak     : BOOL;                      // 开阀确认计时器断输入一拍 / open window one-scan break
    _bCloseBreak  : BOOL;                      // 关阀确认计时器断输入一拍 / close window one-scan break
    _bDrainBreak  : BOOL;                      // 排空计时器断输入一拍 / drain window one-scan break
    _bTotalBreak  : BOOL;                      // 总时长计时器断输入一拍 / total timer one-scan break
    _bVolumeOk    : BOOL;                      // 累计量达目标 / the target volume is reached
    _bRunning     : BOOL;                      // 处于计时阶段（准备/转移/排空/关阀） / inside a timed phase
    _bDrainedHeld : BOOL;                      // 排空完成保持量 / held drained flag
    _bCoastBreak  : BOOL;                      // 惰转计时器断输入一拍 / coast window one-scan break
    _bAbortCloseBreak : BOOL;                  // 中止关阀确认计时器断输入一拍 / abort close window one-scan break
    _bAbortCloseToAcc : BOOL;                  // 中止关阀确认超时锁存（等新启动清除） / held abort close-confirm timeout latch
END_VAR
VAR CONSTANT
    DL_VAL_LIM    : REAL := 1.0E9;             // 有限性判定的绝对值上限 [无量纲] / finiteness ceiling
    DL_VOL_MIN    : REAL := 0.0;               // 目标体积下限 [m3]，须严格大于 / target volume floor, strictly greater
    DL_FLOW_MIN   : REAL := 0.0;               // 排空门限下限 [m3/h] / drain threshold floor [m3/h]
    DL_TIME_ZERO  : TIME := T#0MS;             // 时间零值基准 [ms] / time zero reference
END_VAR

(*------------------------------------------------------------------------------
 * 段 1｜每拍预置：泵与双阀**先全清**（R72），单拍标志预清零（R25 第一律）
 *      Pump and both valves cleared first, one-shot flags pre-cleared
 *-----------------------------------------------------------------------------*)
bPumpCmd     := FALSE;                         // 泵指令先清 / pump command cleared first
bSrcValveCmd := FALSE;                         // 源阀指令先清 / source valve cleared first
bDstValveCmd := FALSE;                         // 目标阀指令先清 / destination valve cleared first
bDrained     := FALSE;                         // 排空标志每拍重算 / drained flag recomputed
bDone        := FALSE;                         // 完成标志每拍重算 / done flag recomputed
bFailed      := FALSE;                         // 失败标志每拍重算 / failed flag recomputed
bValid       := FALSE;                         // 可用标志每拍重算 / usable flag recomputed
eErr         := 16#0000_0000;                  // 错误码每拍重算 / error code recomputed
bError       := FALSE;                         // 故障标志每拍重算 / fault flag recomputed
_bParamBad   := FALSE;                         // 参数非法标志预清零 / parameter flag pre-cleared
_bFiniteBad  := FALSE;                         // 非有限标志预清零 / non-finite flag pre-cleared
_bIllegal    := FALSE;                         // 非法状态标志预清零 / illegal state flag pre-cleared
_bBothFb     := FALSE;                         // 双阀到位标志预置 FALSE / both-feedback preset FALSE
_bDrainCond  := FALSE;                         // 排空条件预置 FALSE / drain condition preset FALSE
_bVolumeOk   := FALSE;                         // 体积达标预置 FALSE / volume reached preset FALSE
_bRunning    := FALSE;                         // 计时阶段标志预置 FALSE / running preset FALSE

(*------------------------------------------------------------------------------
 * 段 2｜首扫初始化（锁存与保持量从零起）
 *      First-scan initialisation
 *-----------------------------------------------------------------------------*)
IF NOT _bInit THEN
    _eState       := E_DL_TransferState.eIdle;  // 相位待机 / phase idle
    _bFaultAcc    := FALSE;                     // 故障锁存清零 / fault latch cleared
    _bFailedAcc   := FALSE;                     // 失败锁存清零 / failure latch cleared
    _bDrainedHeld := FALSE;                     // 排空保持量清零 / drained flag cleared
    _bAbortCloseToAcc := FALSE;                 // 中止关阀确认超时锁存清零 / abort close timeout latch cleared
    _bFbBreak     := TRUE;                      // 开阀确认窗从零开始 / the open window starts from zero
    _bCloseBreak  := TRUE;                      // 关阀确认窗从零开始 / the close window starts from zero
    _bDrainBreak  := TRUE;                      // 排空验证窗从零开始 / the drain window starts from zero
    _bTotalBreak  := TRUE;                      // 总时长计时从零开始 / the total timer starts from zero
    _bInit        := TRUE;                      // 首扫只做一次 / the first scan runs once
END_IF

(*------------------------------------------------------------------------------
 * 段 3｜参数闸门（目标体积、总超时、排空门限）
 *      Parameter gate for the target volume, the timeout and the drain threshold
 *-----------------------------------------------------------------------------*)
IF (fVolumeTarget <> fVolumeTarget) OR (ABS(fVolumeTarget) > DL_VAL_LIM) OR (fVolumeTarget <= DL_VOL_MIN) THEN
    _bParamBad := TRUE;                        // 目标体积非法 / target volume illegal
END_IF
IF TIME_TO_DINT(tTimeout) <= 0 THEN
    _bParamBad := TRUE;                        // 总超时为 0：无限等待，非法 / zero timeout means waiting forever
END_IF
IF xCoastStop AND (TIME_TO_DINT(tPumpCoastTime) <= 0) THEN
    _bParamBad := TRUE;                        // 两段化已使能但惰转窗为 0：退化为单拍中止，违背修复意图，按非法参数拦截 / coast time of zero degrades the two-stage abort, intercepted as an illegal parameter
END_IF
IF (fDrainFlow <> fDrainFlow) OR (ABS(fDrainFlow) > DL_VAL_LIM) OR (fDrainFlow < DL_FLOW_MIN) THEN
    _bParamBad := TRUE;                        // 排空门限非法 / drain threshold illegal
END_IF

(*------------------------------------------------------------------------------
 * 段 4｜输入有限性（累计量与流量；区间判据同时拦 NaN 与 ±Inf）
 *      Input finiteness for the injected volume and the flow
 *-----------------------------------------------------------------------------*)
IF (fTransferred < -DL_VAL_LIM) OR (fTransferred > DL_VAL_LIM) THEN
    _bFiniteBad := TRUE;                       // 累计量非有限 / injected volume non-finite
END_IF
IF (fFlow < -DL_VAL_LIM) OR (fFlow > DL_VAL_LIM) THEN
    _bFiniteBad := TRUE;                       // 流量非有限 / flow non-finite
END_IF

(*------------------------------------------------------------------------------
 * 段 5｜判据计算（双阀到位 / 体积达标 / 排空条件 / 计时阶段）
 *      Criteria evaluation
 *-----------------------------------------------------------------------------*)
_bBothFb    := bSrcValveFb AND bDstValveFb;    // 双阀同时到位（启泵的唯一许可） / both valves open, the only permit to start the pump
_bVolumeOk  := (fTransferred >= fVolumeTarget); // 累计量达目标 [布尔] / the target volume is reached
_bDrainCond := (fFlow < fDrainFlow);           // 排空条件：流量低于门限 / drain condition

_bRunning := (_eState = E_DL_TransferState.ePrepValve)
             OR (_eState = E_DL_TransferState.eTransferring)
             OR (_eState = E_DL_TransferState.eDraining)
             OR (_eState = E_DL_TransferState.eClosing);

(*------------------------------------------------------------------------------
 * 段 6｜四只计时器无条件刷新（R40：CASE 之外每拍必调，各司其职不复用）
 *      Four timers refreshed unconditionally, one duty each, never reused
 *-----------------------------------------------------------------------------*)
fbValveFb(IN := (_eState = E_DL_TransferState.ePrepValve) AND (NOT _bFbBreak), PT := tValveFb); // 开阀到位确认窗
_bFbBreak := FALSE;                            // 断输入拍在调用后自清 / break self-cleared after the call

fbCloseFb(IN := (_eState = E_DL_TransferState.eClosing) AND (NOT _bCloseBreak), PT := tValveFb); // 关阀确认窗
_bCloseBreak := FALSE;                         // 断输入拍在调用后自清 / break self-cleared after the call

fbDrain(IN := (_eState = E_DL_TransferState.eDraining) AND _bDrainCond AND (NOT _bDrainBreak),
        PT := tDrainVerify);                   // 排空验证窗
_bDrainBreak := FALSE;                         // 断输入拍在调用后自清 / break self-cleared after the call

fbTotal(IN := _bRunning AND (NOT _bTotalBreak), PT := tTimeout); // 转移总时长
_bTotalBreak := FALSE;                         // 断输入拍在调用后自清 / break self-cleared after the call

fbCoast(IN := (_eState = E_DL_TransferState.eAbortCoast) AND (NOT _bCoastBreak), PT := tPumpCoastTime); // 泵惰转计时窗（中止第一段）
_bCoastBreak := FALSE;                         // 断输入拍在调用后自清 / break self-cleared after the call

fbAbortClose(IN := (_eState = E_DL_TransferState.eAbortClose) AND (bSrcValveFb OR bDstValveFb) AND (NOT _bAbortCloseBreak),
             PT := tValveFb);                  // 中止关阀确认窗：阀开反馈任一保持即计时 / abort close window, timed while any open feedback holds
_bAbortCloseBreak := FALSE;                    // 断输入拍在调用后自清 / break self-cleared after the call

(*------------------------------------------------------------------------------
 * 段 7｜相位机（只做迁移；输出在段 8 按相置位，泵永远在阀之后）
 *      Phase machine, transitions only, the pump is always gated behind the valves
 *-----------------------------------------------------------------------------*)
IF bAbort AND (_eState <> E_DL_TransferState.eAbort)
   AND (_eState <> E_DL_TransferState.eAbortCoast) AND (_eState <> E_DL_TransferState.eAbortClose) THEN
    (* 中止：任意拍生效；中止族态内不重复触发（防惰转窗被反复重启，v1.0.2） *)
    (* Abort takes effect on any scan, not re-triggered inside the abort family *)
    IF xCoastStop THEN
        _eState    := E_DL_TransferState.eAbortCoast; // 两段化：先断泵、阀保持，惰转计时 / two-stage: pump off, valves held, coast timing
        _bCoastBreak := TRUE;                  // 惰转窗从零开始 / the coast window starts from zero
    ELSE
        _eState    := E_DL_TransferState.eAbort; // 兼容路径：单拍停泵关阀（不推荐） / legacy single-scan abort, not recommended
    END_IF
    _bFbBreak  := TRUE;                        // 四个窗全部重启 / every window restarts
    _bCloseBreak := TRUE;
    _bDrainBreak := TRUE;
    _bTotalBreak := TRUE;
    _bAbortCloseBreak := TRUE;                 // 中止关阀确认窗重启 / the abort close window restarts
ELSIF _bParamBad THEN
    _eState := E_DL_TransferState.eFault;      // 参数非法：转故障 / illegal parameters go to fault
    _bFailedAcc := TRUE;                       // 失败锁存（本批不可用） / this batch is unusable
ELSIF _bFiniteBad THEN
    _eState := E_DL_TransferState.eFault;      // 输入非有限：转故障，停泵关阀（段 8） / non-finite input
    _bFailedAcc := TRUE;                       // 失败锁存 / failure latched
ELSE
    IF fbTotal.Q AND _bRunning THEN
        (* 总时长超时：先锁存失败再转故障，段 8 下一拍停泵关阀 *)
        (* Total timeout, the failure is latched and the outputs drop on the next scan *)
        _bFailedAcc := TRUE;                   // 本批失败锁定 / latch the failure
        _bFbBreak   := TRUE;                   // 四个窗全部重启 / every window restarts
        _bCloseBreak := TRUE;
        _bDrainBreak := TRUE;
        _bTotalBreak := TRUE;
        _eState     := E_DL_TransferState.eFault;
    ELSIF (_eState <> E_DL_TransferState.eIdle) AND (_eState <> E_DL_TransferState.eAbort)
          AND (_eState <> E_DL_TransferState.eAbortCoast) AND (_eState <> E_DL_TransferState.eAbortClose)
          AND (_eState <> E_DL_TransferState.eFault) AND (NOT bStart) THEN
        (* 启动撤销等同中止：外部撤掉启动必须让设备停下，不能继续跑 *)
        (* A dropped start is treated as an abort, the machine must stop *)
        IF xCoastStop THEN
            _eState      := E_DL_TransferState.eAbortCoast; // 两段化中止 / two-stage abort
            _bCoastBreak := TRUE;               // 惰转窗从零开始 / the coast window starts from zero
        ELSE
            _eState      := E_DL_TransferState.eAbort; // 兼容路径单拍中止 / legacy single-scan abort
        END_IF
        _bFbBreak  := TRUE;
        _bCloseBreak := TRUE;
        _bDrainBreak := TRUE;
        _bTotalBreak := TRUE;
        _bAbortCloseBreak := TRUE;              // 中止关阀确认窗重启 / the abort close window restarts
    ELSE
        CASE _eState OF

            E_DL_TransferState.eIdle:          // 待机：启动即准备阀门
                IF bStart THEN
                    _bFaultAcc    := FALSE;    // 新任务清除故障锁存 / a new job clears the fault latch
                    _bFailedAcc   := FALSE;    // 新任务清除失败锁存 / a new job clears the failure latch
                    _bDrainedHeld := FALSE;    // 新任务清除排空保持量 / a new job clears the drained flag
                    _bAbortCloseToAcc := FALSE; // 新任务清除中止关阀超时锁存 / a new job clears the abort close timeout latch
                    _bFbBreak     := TRUE;     // 开阀确认窗从零开始 / the open window starts from zero
                    _bTotalBreak  := TRUE;     // 总时长从零开始 / the total timer starts from zero
                    _eState       := E_DL_TransferState.ePrepValve; // 进准备阀门相 / prepare the valves
                END_IF

            E_DL_TransferState.ePrepValve:     // 准备阀门：双阀到位才启泵
                IF _bBothFb THEN
                    _bTotalBreak := TRUE;      // 启泵当拍重启总时长（此前只算阀门准备） / the total timer restarts at pump start
                    _eState      := E_DL_TransferState.eTransferring; // 进转移相 / start transferring
                ELSIF fbValveFb.Q THEN
                    _bFaultAcc := TRUE;        // 阀位反馈超时：锁存故障 / feedback timeout, latch the fault
                    _bFbBreak  := TRUE;        // 窗重启 / the window restarts
                    _eState    := E_DL_TransferState.eIdle; // 回待机（先清输出，泵从未启动） / back to idle
                END_IF

            E_DL_TransferState.eTransferring:  // 转移中：累计量达目标即停泵
                IF _bVolumeOk THEN
                    _bDrainBreak := TRUE;      // 排空验证窗从零开始 / the drain window starts from zero
                    _eState      := E_DL_TransferState.eDraining; // 进排空相（泵在段 8 停） / start draining
                END_IF

            E_DL_TransferState.eDraining:      // 排空中：流量持续低于门限即判排空完成
                IF fbDrain.Q THEN
                    _bDrainedHeld := TRUE;     // 排空完成（保持量） / drained, latched
                    _bCloseBreak  := TRUE;     // 关阀确认窗从零开始 / the close window starts from zero
                    _eState       := E_DL_TransferState.eClosing; // 进关阀相 / close the valves
                END_IF

            E_DL_TransferState.eClosing:       // 关阀中：确认窗满即完成
                IF fbCloseFb.Q THEN
                    _eState := E_DL_TransferState.eComplete; // 进完成相 / complete
                END_IF

            E_DL_TransferState.eComplete:      // 完成：等启动撤销（bStart 落下由上方统一处理）
                _bTotalBreak := TRUE;          // 总时长停表 / stop the total timer
                _bFbBreak    := TRUE;          // 各窗复位 / every window reset
                _bCloseBreak := TRUE;
                _bDrainBreak := TRUE;

            E_DL_TransferState.eAbort:         // 中止兼容路径：等启动撤销后回待机
                _bTotalBreak := TRUE;          // 总时长停表 / stop the total timer
                IF NOT bStart THEN
                    _eState := E_DL_TransferState.eIdle; // 启动已撤销，回待机 / back to idle
                END_IF

            E_DL_TransferState.eAbortCoast:    // 中止第一段：泵已断使能、阀保持不动，等惰转窗满
                _bTotalBreak := TRUE;          // 总时长停表 / stop the total timer
                IF fbCoast.Q THEN
                    _bAbortCloseBreak := TRUE; // 惰转窗满，中止关阀确认窗从零开始 / coast elapsed, the abort close window starts from zero
                    _eState := E_DL_TransferState.eAbortClose; // 进中止第二段（阀指令在段 8 清零）/ abort stage B
                END_IF

            E_DL_TransferState.eAbortClose:    // 中止第二段：关阀指令已发，等阀离开开位或确认超时
                _bTotalBreak := TRUE;          // 总时长停表 / stop the total timer
                IF fbAbortClose.Q THEN
                    _bAbortCloseToAcc := TRUE; // 阀开反馈在确认窗内保持：关阀确认超时锁存 / open feedback held through the window, close-confirm timeout latched
                END_IF
                IF (NOT bSrcValveFb) AND (NOT bDstValveFb) AND (NOT bStart) THEN
                    _eState := E_DL_TransferState.eIdle; // 阀已离开开位且启动撤销，回待机 / valves left open position and the start is dropped
                END_IF

            E_DL_TransferState.eFault:         // 故障：启动撤销且参数合法才回待机
                IF (NOT bStart) AND (NOT _bParamBad) AND (NOT _bFiniteBad) THEN
                    _eState := E_DL_TransferState.eIdle; // 原因消失 / the cause is gone
                END_IF

            ELSE
                _bIllegal := TRUE;             // 标记非法状态 / flag the illegal state
                _bFbBreak := TRUE;             // 四个窗全部重启 / every window restarts
                _bCloseBreak := TRUE;
                _bDrainBreak := TRUE;
                _bTotalBreak := TRUE;
                _eState := E_DL_TransferState.eFault; // 回故障态 / back to the fault state
        END_CASE
    END_IF
END_IF

(*------------------------------------------------------------------------------
 * 段 8｜输出置位（次序即安全：**泵先于阀**，中止路径先停泵后关阀）
 *      Output assignment, the pump always precedes the valves
 *-----------------------------------------------------------------------------*)
CASE _eState OF
    E_DL_TransferState.ePrepValve:             // 准备阀门：双阀开，泵不启
        bSrcValveCmd := TRUE;                  // 源阀开 / source valve open
        bDstValveCmd := TRUE;                  // 目标阀开 / destination valve open
    E_DL_TransferState.eTransferring:          // 转移：双阀保持 + 泵运行（泵在阀之后赋值）
        bSrcValveCmd := TRUE;                  // 源阀开 / source valve open
        bDstValveCmd := TRUE;                  // 目标阀开 / destination valve open
        bPumpCmd     := TRUE;                  // 泵运行（阀门已到位并保持） / the pump runs after the valves are open
    E_DL_TransferState.eDraining:              // 排空：泵停、双阀仍开
        bSrcValveCmd := TRUE;                  // 源阀开 / source valve open
        bDstValveCmd := TRUE;                  // 目标阀开 / destination valve open
    E_DL_TransferState.eAbortCoast:            // 中止第一段：泵断使能、**阀位保持不动**（不发关阀指令，
                                               //   机检断言：abort 拍不得出现关阀输出置位，验收向量 V9/V10）
        bSrcValveCmd := TRUE;                  // 源阀保持开（惰转窗内阀位不动） / source valve held open during the coast window
        bDstValveCmd := TRUE;                  // 目标阀保持开 / destination valve held open
    ELSE
        bPumpCmd     := FALSE;                 // 其余相：泵显式停（先停泵） / pump explicitly stopped first
        bSrcValveCmd := FALSE;                 // 源阀关指令（TRUE = 开启，故清指令即关阀） / source valve closed
        bDstValveCmd := FALSE;                 // 目标阀关指令 / destination valve closed
END_CASE

(*------------------------------------------------------------------------------
 * 段 9｜码位优先级链与出口
 *      Code priority chain and exit
 *-----------------------------------------------------------------------------*)
IF _bIllegal THEN
    eErr     := 16#0005_0316;                  // 故障级：状态机兜底 / fault: state machine fallback
    bError   := TRUE;                          // 置故障标志 / raise the fault flag
    _bFailedAcc := TRUE;                       // 非法状态按失败锁定 / an illegal state latches a failure
ELSIF _bParamBad OR _bFiniteBad THEN
    eErr     := 16#0005_0315;                  // 故障级：参数非法或输入非有限（复用，R90） / fault: illegal parameter or non-finite input
    bError   := TRUE;                          // 置故障标志 / raise the fault flag
ELSIF _bAbortCloseToAcc THEN
    eErr     := 16#0005_0317;                  // 故障级：中止第二段关阀确认超时（v1.0.2 新增） / fault: abort close-confirm timeout
    bError   := TRUE;                          // 故障级码位必须同时置故障标志（R45 配对） / a fault-class code must raise the fault flag
ELSIF (_eState = E_DL_TransferState.eFault) AND _bFailedAcc THEN
    eErr     := 16#0005_0315;                  // 故障级：转移总时长超时（复用，R90） / fault: total transfer timeout
    bError   := TRUE;                          // 故障级码位必须置故障标志（R22 终审修复：原实现漏置）/ a fault-class code must raise the fault flag
ELSIF _bFaultAcc THEN
    eErr     := 16#0005_0314;                  // 故障级：阀位反馈超时未到位，拒绝启泵 / fault: feedback timeout, no pump start
    bError   := TRUE;                          // 置故障标志 / raise the fault flag
ELSIF _bDrainedHeld THEN
    eErr     := 16#0005_01E1;                  // 信息级：排空验证窗内流量持续低于门限 / informational: drained
ELSIF _eState = E_DL_TransferState.eTransferring THEN
    eErr     := 16#0005_01E0;                  // 信息级：累计量由调用方注入，本件不重复积分 / informational: the volume is injected
END_IF

bDrained   := _bDrainedHeld;                   // 排空标志出口 / drained outlet
bDone      := (_eState = E_DL_TransferState.eComplete); // 完成放行出口 / done outlet
bFailed    := (_eState = E_DL_TransferState.eFault) OR _bFailedAcc OR _bAbortCloseToAcc; // 失败出口（中止本身是人的决定不计失败；关阀确认超时是真实故障，计入）

IF bError THEN
    bValid := FALSE;                           // 故障级：输出不可用 / fault: outputs unusable
ELSIF (_eState = E_DL_TransferState.eIdle) THEN
    bValid := FALSE;                           // 待机：无批次在执行 / idle: no batch in progress
ELSE
    bValid := TRUE;                            // 输出可用 / outputs usable
END_IF

END_FUNCTION_BLOCK
